(* IEC 61131-3 sources: plc-st-coding-agent/progress/evidence/f14_v10_full_20261113/jobs/custom_minimax-m27 (part 8) *)

(* ---- self-medium-01.candidate_03.st ---- *)
(* ENGINEERING_CONTRACT *)
(*
  PUB002/PUB005: valid=FALSE → loadedID:=0, valid=TRUE → loadedID:=recipe[selSlot].recipeID
  PUB006: loadCmd rising-edge triggers one-shot load; level-hold does NOT reload
  PUB007: running=TRUE blocks load, loadedID retains previous value
  PUB008: slot out-of-range [1..8] → valid=FALSE, loadedID unchanged; no array OOB access
  PUB009: validation is conjunction: recipeID<>0 AND totalRatio∈[99.0,101.0] AND temperature∈[30.0,180.0]
  Timing: state retention via VAR (static across scans); first-scan prev_* = FALSE (IEC default)
  S1: !running & rising(loadCmd) & valid-slot & empty-slot → valid=FALSE & loadedID=0
  S4/N10-S4: running → loadedID=prev(loadedID) (includes first production entry)
  N10-S9: !running & !rising(loadCmd) → both outputs retain prev value
*)
(* CONTRACT_RULES [] *)

FUNCTION_BLOCK FB
VAR_INPUT
    recipe      : ARRAY[1..8] OF ST_Recipe;
    selSlot     : INT;
    loadCmd     : BOOL;
    running     : BOOL;
END_VAR
VAR_OUTPUT
    valid       : BOOL;
    loadedID    : INT;
END_VAR
VAR
    tmp_loadTrig  : R_TRIG;
    tmp_prevRunning : BOOL := FALSE;
END_VAR

tmp_loadTrig(CLK := loadCmd);

IF tmp_loadTrig.Q AND NOT running THEN
    IF (selSlot >= 1) AND (selSlot <= 8) THEN
        IF (recipe[selSlot].recipeID <> 0) AND
           (recipe[selSlot].totalRatio >= 99.0) AND (recipe[selSlot].totalRatio <= 101.0) AND
           (recipe[selSlot].temperature >= 30.0) AND (recipe[selSlot].temperature <= 180.0) THEN
            valid    := TRUE;
            loadedID := recipe[selSlot].recipeID;
        ELSE
            valid    := FALSE;
            loadedID := 0;
        END_IF;
    ELSE
        valid    := FALSE;
    END_IF;
ELSIF running THEN
    loadedID := loadedID;
END_IF;

tmp_prevRunning := running;
END_FUNCTION_BLOCK

(* ---- self-medium-01.raw_candidate_01.st ---- *)
(* ENGINEERING_CONTRACT *)
(*
  PUB002/PUB005: valid=FALSE → loadedID:=0, valid=TRUE → loadedID:=recipe[selSlot].recipeID
  PUB006: loadCmd rising-edge triggers one-shot load; level-hold does NOT reload
  PUB007: running=TRUE blocks load, loadedID retains previous value
  PUB008: slot out-of-range [1..8] → valid=FALSE, loadedID unchanged; no array OOB access
  PUB009: validation is conjunction: recipeID<>0 AND totalRatio∈[99.0,101.0] AND temperature∈[30.0,180.0]
  Timing: state retention via VAR (static across scans); first-scan prev_* = FALSE (IEC default)
  S1: !running & rising(loadCmd) & valid-slot & empty-slot → valid=FALSE & loadedID=0
  S4/N10-S4: running → loadedID=prev(loadedID) (includes first production entry)
  N10-S9: !running & !rising(loadCmd) → both outputs retain prev value
*)
(* CONTRACT_RULES [] *)

FUNCTION_BLOCK FB
VAR_INPUT
    recipe      : ARRAY[1..8] OF ST_Recipe;
    selSlot     : INT;
    loadCmd     : BOOL;
    running     : BOOL;
END_VAR
VAR_OUTPUT
    valid       : BOOL;
    loadedID    : INT;
END_VAR
VAR
    tmp_loadTrig  : R_TRIG;
    tmp_prevRunning : BOOL := FALSE;
END_VAR

tmp_loadTrig(CLK := loadCmd);

IF tmp_loadTrig.Q AND NOT running THEN
    IF (selSlot >= 1) AND (selSlot <= 8) THEN
        IF (recipe[selSlot].recipeID <> 0) AND
           (recipe[selSlot].totalRatio >= 99.0) AND (recipe[selSlot].totalRatio <= 101.0) AND
           (recipe[selSlot].temperature >= 30.0) AND (recipe[selSlot].temperature <= 180.0) THEN
            valid    := TRUE;
            loadedID := recipe[selSlot].recipeID;
        ELSE
            valid    := FALSE;
            loadedID := 0;
        END_IF;
    ELSE
        valid    := FALSE;
    END_IF;
ELSIF running THEN
    loadedID := loadedID;
END_IF;

tmp_prevRunning := running;

(* ---- self-medium-01.raw_candidate_02.st ---- *)
(* ENGINEERING_CONTRACT *)
(*
  PUB002/PUB005: valid=FALSE → loadedID:=0, valid=TRUE → loadedID:=recipe[selSlot].recipeID
  PUB006: loadCmd rising-edge triggers one-shot load; level-hold does NOT reload
  PUB007: running=TRUE blocks load, loadedID retains previous value
  PUB008: slot out-of-range [1..8] → valid=FALSE, loadedID unchanged; no array OOB access
  PUB009: validation is conjunction: recipeID<>0 AND totalRatio∈[99.0,101.0] AND temperature∈[30.0,180.0]
  Timing: state retention via VAR (static across scans); first-scan prev_* = FALSE (IEC default)
  S1: !running & rising(loadCmd) & valid-slot & empty-slot → valid=FALSE & loadedID=0
  S4/N10-S4: running → loadedID=prev(loadedID) (includes first production entry)
  N10-S9: !running & !rising(loadCmd) → both outputs retain prev value
*)
(* CONTRACT_RULES [] *)

FUNCTION_BLOCK FB
VAR_INPUT
    recipe      : ARRAY[1..8] OF ST_Recipe;
    selSlot     : INT;
    loadCmd     : BOOL;
    running     : BOOL;
END_VAR
VAR_OUTPUT
    valid       : BOOL;
    loadedID    : INT;
END_VAR
VAR
    tmp_loadTrig  : R_TRIG;
    tmp_prevRunning : BOOL := FALSE;
END_VAR

tmp_loadTrig(CLK := loadCmd);

IF tmp_loadTrig.Q AND NOT running THEN
    IF (selSlot >= 1) AND (selSlot <= 8) THEN
        IF (recipe[selSlot].recipeID <> 0) AND
           (recipe[selSlot].totalRatio >= 99.0) AND (recipe[selSlot].totalRatio <= 101.0) AND
           (recipe[selSlot].temperature >= 30.0) AND (recipe[selSlot].temperature <= 180.0) THEN
            valid    := TRUE;
            loadedID := recipe[selSlot].recipeID;
        ELSE
            valid    := FALSE;
            loadedID := 0;
        END_IF;
    ELSE
        valid    := FALSE;
    END_IF;
ELSIF running THEN
    loadedID := loadedID;
END_IF;

tmp_prevRunning := running;
END_FUNCTION_BLOCK

(* ---- self-medium-01.raw_candidate_03.st ---- *)
(* ENGINEERING_CONTRACT *)
(*
  PUB002/PUB005: valid=FALSE → loadedID:=0, valid=TRUE → loadedID:=recipe[selSlot].recipeID
  PUB006: loadCmd rising-edge triggers one-shot load; level-hold does NOT reload
  PUB007: running=TRUE blocks load, loadedID retains previous value
  PUB008: slot out-of-range [1..8] → valid=FALSE, loadedID unchanged; no array OOB access
  PUB009: validation is conjunction: recipeID<>0 AND totalRatio∈[99.0,101.0] AND temperature∈[30.0,180.0]
  Timing: state retention via VAR (static across scans); first-scan prev_* = FALSE (IEC default)
  S1: !running & rising(loadCmd) & valid-slot & empty-slot → valid=FALSE & loadedID=0
  S4/N10-S4: running → loadedID=prev(loadedID) (includes first production entry)
  N10-S9: !running & !rising(loadCmd) → both outputs retain prev value
*)
(* CONTRACT_RULES [] *)

FUNCTION_BLOCK FB
VAR_INPUT
    recipe      : ARRAY[1..8] OF ST_Recipe;
    selSlot     : INT;
    loadCmd     : BOOL;
    running     : BOOL;
END_VAR
VAR_OUTPUT
    valid       : BOOL;
    loadedID    : INT;
END_VAR
VAR
    tmp_loadTrig  : R_TRIG;
    tmp_prevRunning : BOOL := FALSE;
END_VAR

tmp_loadTrig(CLK := loadCmd);

IF tmp_loadTrig.Q AND NOT running THEN
    IF (selSlot >= 1) AND (selSlot <= 8) THEN
        IF (recipe[selSlot].recipeID <> 0) AND
           (recipe[selSlot].totalRatio >= 99.0) AND (recipe[selSlot].totalRatio <= 101.0) AND
           (recipe[selSlot].temperature >= 30.0) AND (recipe[selSlot].temperature <= 180.0) THEN
            valid    := TRUE;
            loadedID := recipe[selSlot].recipeID;
        ELSE
            valid    := FALSE;
            loadedID := 0;
        END_IF;
    ELSE
        valid    := FALSE;
    END_IF;
ELSIF running THEN
    loadedID := loadedID;
END_IF;

tmp_prevRunning := running;
END_FUNCTION_BLOCK

(* ---- self-medium-02.candidate_01.st ---- *)
FUNCTION_BLOCK FB
VAR_INPUT
    enable     : BOOL;
    rawValue   : REAL;
END_VAR
VAR_OUTPUT
    filteredValue : REAL;
    windowFull    : BOOL;
    sampleCount   : INT;
END_VAR
VAR
    buffer     : ARRAY[0..7] OF REAL;
    writeIdx   : INT := 0;
    tmp_sum    : REAL;
    tmp_i      : INT;
END_VAR
VAR_INPUT
END_VAR
VAR_OUTPUT
END_VAR
VAR
END_VAR
(* ENGINEERING_CONTRACT
   PUB.001-004   : inputs enable, rawValue; outputs filteredValue, windowFull, sampleCount
   PUB.005       : enable=TRUE per scan: push rawValue into 8-slot ring buffer
   PUB.006       : filteredValue = mean of actually-filled slots (no zero-fill)
   PUB.007       : on windowFull: FIFO eviction of oldest sample on each new push
   PUB.008       : sampleCount = current valid samples 0..8
   PUB.009       : windowFull = TRUE when sampleCount == 8, retains TRUE thereafter
   PUB.010       : enable=FALSE: clear buffer (sampleCount=0, windowFull=FALSE),
                   filteredValue RETAINED (last computed value held)
   PUB.011       : new enable period restarts count from 1 independently
   PUB.012-015   : formal properties S1-S7 encoded as LTL constraints
   PUB.016-038   : interface unchanged; no hidden timers or global variables

   Output retention table:
   | output        | activation             | retention      | reset                    |
   |---------------|------------------------|----------------|--------------------------|
   | filteredValue | every enabled scan     | holds on FALSE | not reset; retains last  |
   | sampleCount   | increments on each push| capped at 8    | forced 0 on enable=FALSE |
   | windowFull    | set TRUE at count=8    | holds TRUE     | forced FALSE on enable=FALSE|

   Same-scan priority: disable branch executes first; rising-edge start is
   indistinguishable from normal enabled scan since buffer is pre-cleared.
   Units: filteredValue REAL; sampleCount INT 0..8; windowFull BOOL.

   CONTRACT_RULES []
*)
tmp_sum := 0.0;
IF NOT enable THEN
    sampleCount   := 0;
    windowFull    := FALSE;
    writeIdx      := 0;
ELSE
    // Push current rawValue into ring buffer
    buffer[writeIdx] := rawValue;

    // Advance write pointer (mod 8), but sampleCount only increments up to 8
    writeIdx := (writeIdx + 1) MOD 8;
    IF sampleCount < 8 THEN
        sampleCount := sampleCount + 1;
    END_IF;

    // windowFull stays TRUE once set; set it only when count reaches 8
    IF sampleCount = 8 THEN
        windowFull := TRUE;
    END_IF;

    // Compute arithmetic mean of all valid samples currently in buffer
    tmp_sum := 0.0;
    FOR tmp_i := 0 TO sampleCount - 1 DO
        tmp_sum := tmp_sum + buffer[tmp_i];
    END_FOR;
    filteredValue := tmp_sum / TO_REAL(sampleCount);
END_IF;
END_FUNCTION_BLOCK

(* ---- self-medium-02.raw_candidate_01.st ---- *)
FUNCTION_BLOCK FB
VAR_INPUT
    enable     : BOOL;
    rawValue   : REAL;
END_VAR
VAR_OUTPUT
    filteredValue : REAL;
    windowFull    : BOOL;
    sampleCount   : INT;
END_VAR
VAR
    buffer     : ARRAY[0..7] OF REAL;
    writeIdx   : INT := 0;
    tmp_sum    : REAL;
    tmp_i      : INT;
END_VAR
VAR_INPUT
END_VAR
VAR_OUTPUT
END_VAR
VAR
END_VAR
(* ENGINEERING_CONTRACT
   PUB.001-004   : inputs enable, rawValue; outputs filteredValue, windowFull, sampleCount
   PUB.005       : enable=TRUE per scan: push rawValue into 8-slot ring buffer
   PUB.006       : filteredValue = mean of actually-filled slots (no zero-fill)
   PUB.007       : on windowFull: FIFO eviction of oldest sample on each new push
   PUB.008       : sampleCount = current valid samples 0..8
   PUB.009       : windowFull = TRUE when sampleCount == 8, retains TRUE thereafter
   PUB.010       : enable=FALSE: clear buffer (sampleCount=0, windowFull=FALSE),
                   filteredValue RETAINED (last computed value held)
   PUB.011       : new enable period restarts count from 1 independently
   PUB.012-015   : formal properties S1-S7 encoded as LTL constraints
   PUB.016-038   : interface unchanged; no hidden timers or global variables

   Output retention table:
   | output        | activation             | retention      | reset                    |
   |---------------|------------------------|----------------|--------------------------|
   | filteredValue | every enabled scan     | holds on FALSE | not reset; retains last  |
   | sampleCount   | increments on each push| capped at 8    | forced 0 on enable=FALSE |
   | windowFull    | set TRUE at count=8    | holds TRUE     | forced FALSE on enable=FALSE|

   Same-scan priority: disable branch executes first; rising-edge start is
   indistinguishable from normal enabled scan since buffer is pre-cleared.
   Units: filteredValue REAL; sampleCount INT 0..8; windowFull BOOL.

   CONTRACT_RULES []
*)
tmp_sum := 0.0;
IF NOT enable THEN
    sampleCount   := 0;
    windowFull    := FALSE;
    writeIdx      := 0;
ELSE
    // Push current rawValue into ring buffer
    buffer[writeIdx] := rawValue;

    // Advance write pointer (mod 8), but sampleCount only increments up to 8
    writeIdx := (writeIdx + 1) MOD 8;
    IF sampleCount < 8 THEN
        sampleCount := sampleCount + 1;
    END_IF;

    // windowFull stays TRUE once set; set it only when count reaches 8
    IF sampleCount = 8 THEN
        windowFull := TRUE;
    END_IF;

    // Compute arithmetic mean of all valid samples currently in buffer
    tmp_sum := 0.0;
    FOR tmp_i := 0 TO sampleCount - 1 DO
        tmp_sum := tmp_sum + buffer[tmp_i];
    END_FOR;
    filteredValue := tmp_sum / TO_REAL(sampleCount);
END_IF;
END_FUNCTION_BLOCK

(* ---- self-medium-03.candidate_01.st ---- *)
(* ENGINEERING_CONTRACT *)
(*
  Gate FSM: 4 states (IDLE/OPENING/CLOSING/FAULT), obstacle safety interlock.

  PUB001: IDLE at power-on, initial button values FALSE.
  PUB003: Rising edge of openBtn (closeBtn=FALSE, openLimit=FALSE) starts opening.
          Rising edge of closeBtn (openBtn=FALSE, closeLimit=FALSE) starts closing.
          Both buttons simultaneous → no start. Commands issued same scan.
  PUB004: Buttons ignored during OPENING/CLOSING.
  PUB005: At own-direction limit → stop that direction, return IDLE.
          Opposite limit does not affect current motion.
  PUB006: MotorUp and motorDown always mutually exclusive.
  PUB007: Obstacle at any time → stop both motors, enter FAULT, errorFlag:=TRUE immediately.
          Obstacle priority > limit/motion/reset.
  PUB008: FAULT latches errorFlag, stops motors.
  PUB009: Clear fault only when: no obstacle AND both buttons new rising edge from
          not-both-pressed state to both-pressed state. Holding both with obstacle
          present does NOT clear on obstacle-clear scan. Reset→IDLE, both motors stop
          that scan, then normal PUB003 rules apply.
*)
TYPE GateState :
(
    IDLE    := 0,
    OPENING := 1,
    CLOSING := 2,
    FAULT   := 3
);
END_TYPE;

FUNCTION_BLOCK FB
VAR_INPUT
    openBtn    : BOOL;
    closeBtn   : BOOL;
    openLimit  : BOOL;
    closeLimit : BOOL;
    obstacle   : BOOL;
END_VAR

VAR_OUTPUT
    motorUp    : BOOL;
    motorDown  : BOOL;
    errorFlag  : BOOL;
END_VAR

VAR
    state        : GateState := IDLE;
    prevOpenBtn  : BOOL := FALSE;
    prevCloseBtn : BOOL := FALSE;
    prevObstacle : BOOL := FALSE;
    prevMotorUp  : BOOL := FALSE;
    prevMotorDown: BOOL := FALSE;
    prevErrorFlag: BOOL := FALSE;
END_VAR

VAR
    risingOpen  : BOOL;
    risingClose : BOOL;
    risingBoth  : BOOL;
END_VAR
(* ENGINEERING_CONTRACT *)
(*
  Gate FSM: 4 states (IDLE/OPENING/CLOSING/FAULT), obstacle safety interlock.

  PUB001: IDLE at power-on, initial button values FALSE.
  PUB003: Rising edge of openBtn (closeBtn=FALSE, openLimit=FALSE) starts opening.
          Rising edge of closeBtn (openBtn=FALSE, closeLimit=FALSE) starts closing.
          Both buttons simultaneous → no start. Commands issued same scan.
  PUB004: Buttons ignored during OPENING/CLOSING.
  PUB005: At own-direction limit → stop that direction, return IDLE.
          Opposite limit does not affect current motion.
  PUB006: MotorUp and motorDown always mutually exclusive.
  PUB007: Obstacle at any time → stop both motors, enter FAULT, errorFlag:=TRUE immediately.
          Obstacle priority > limit/motion/reset.
  PUB008: FAULT latches errorFlag, stops motors.
  PUB009: Clear fault only when: no obstacle AND both buttons new rising edge from
          not-both-pressed state to both-pressed state. Holding both with obstacle
          present does NOT clear on obstacle-clear scan. Reset→IDLE, both motors stop
          that scan, then normal PUB003 rules apply.
*)

risingOpen  := openBtn  AND NOT prevOpenBtn;
risingClose := closeBtn AND NOT prevCloseBtn;
risingBoth  := risingOpen AND risingClose;

IF obstacle THEN
    errorFlag  := TRUE;
    motorUp    := FALSE;
    motorDown  := FALSE;
    state      := FAULT;
    GOTO update_state;
END_IF;

IF state = FAULT THEN
    motorUp   := FALSE;
    motorDown := FALSE;
    IF risingBoth THEN
        errorFlag := FALSE;
        state     := IDLE;
    END_IF;
    GOTO update_state;
END_IF;

IF state = IDLE THEN
    IF risingOpen AND NOT closeBtn AND NOT openLimit THEN
        state := OPENING;
    ELSIF risingClose AND NOT openBtn AND NOT closeLimit THEN
        state := CLOSING;
    END_IF;
END_IF;

IF state = OPENING THEN
    motorUp   := TRUE;
    motorDown := FALSE;
    IF openLimit THEN
        motorUp := FALSE;
        state   := IDLE;
    END_IF;
END_IF;

IF state = CLOSING THEN
    motorUp   := FALSE;
    motorDown := TRUE;
    IF closeLimit THEN
        motorDown := FALSE;
        state     := IDLE;
    END_IF;
END_IF;

update_state:
prevOpenBtn   := openBtn;
prevCloseBtn  := closeBtn;
prevObstacle  := obstacle;
prevMotorUp   := motorUp;
prevMotorDown := motorDown;
prevErrorFlag := errorFlag;
END_FUNCTION_BLOCK
(* CONTRACT_RULES [] *)

(* ---- self-medium-03.candidate_02.st ---- *)
(* ENGINEERING_CONTRACT *)
(*
  Gate FSM: 4 states (IDLE/OPENING/CLOSING/FAULT), obstacle safety interlock.
  Priority order (highest first):
  1. Obstacle → stop both, enter FAULT, set errorFlag (same scan).
  2. FAULT → motors held FALSE; reset only on risingBoth when !obstacle.
  3. OPENING/CLOSING → motors set by state; own-limit stops and returns IDLE.
  4. IDLE → rising edge start on single valid button; simultaneous → no start.
  Motors always mutually exclusive (only one direction active at a time).
  Latched outputs: errorFlag (hold_until_reset via risingBoth).
*)
TYPE GateState :
(
    IDLE    := 0,
    OPENING := 1,
    CLOSING := 2,
    FAULT   := 3
);
END_TYPE;

FUNCTION_BLOCK FB
VAR_INPUT
    openBtn    : BOOL;
    closeBtn   : BOOL;
    openLimit  : BOOL;
    closeLimit : BOOL;
    obstacle   : BOOL;
END_VAR

VAR_OUTPUT
    motorUp    : BOOL;
    motorDown  : BOOL;
    errorFlag  : BOOL;
END_VAR

VAR
    state         : GateState := IDLE;
    prevOpenBtn   : BOOL := FALSE;
    prevCloseBtn  : BOOL := FALSE;
    prevMotorUp   : BOOL := FALSE;
    prevMotorDown : BOOL := FALSE;
    prevErrorFlag : BOOL := FALSE;
END_VAR

VAR
    risingOpen  : BOOL;
    risingClose : BOOL;
    risingBoth  : BOOL;
END_VAR

risingOpen  := openBtn  AND NOT prevOpenBtn;
risingClose := closeBtn AND NOT prevCloseBtn;
risingBoth  := openBtn AND closeBtn AND NOT prevOpenBtn AND NOT prevCloseBtn;

IF obstacle THEN
    motorUp   := FALSE;
    motorDown := FALSE;
    errorFlag := TRUE;
    state     := FAULT;
ELSE
    errorFlag := FALSE;

    IF state = FAULT THEN
        motorUp   := FALSE;
        motorDown := FALSE;
        IF risingBoth THEN
            state := IDLE;
        END_IF;

    ELSIF state = IDLE THEN
        motorUp   := FALSE;
        motorDown := FALSE;
        IF risingOpen AND NOT closeBtn AND NOT openLimit THEN
            state := OPENING;
        ELSIF risingClose AND NOT openBtn AND NOT closeLimit THEN
            state := CLOSING;
        END_IF;

    ELSIF state = OPENING THEN
        motorUp   := TRUE;
        motorDown := FALSE;
        IF openLimit THEN
            motorUp := FALSE;
            state   := IDLE;
        END_IF;

    ELSIF state = CLOSING THEN
        motorUp   := FALSE;
        motorDown := TRUE;
        IF closeLimit THEN
            motorDown := FALSE;
            state     := IDLE;
        END_IF;
    END_IF;
END_IF;

prevOpenBtn   := openBtn;
prevCloseBtn  := closeBtn;
prevMotorUp   := motorUp;
prevMotorDown := motorDown;
prevErrorFlag := errorFlag;
END_FUNCTION_BLOCK
(* CONTRACT_RULES [] *)

(* ---- self-medium-03.candidate_03.st ---- *)
Looking at the functional failures, the issue is clear from the replay: `motorUp` is not being set in the same scan as the rising edge triggers the state transition. The motor assignments need to occur after all state transitions, not interleaved within each branch.

```st
(* ENGINEERING_CONTRACT *)
(*
  Gate FSM: 4 states (IDLE/OPENING/CLOSING/FAULT), obstacle safety interlock.
  Priority order (highest first):
  1. Obstacle → stop both, enter FAULT, set errorFlag (same scan).
  2. FAULT → motors held FALSE; reset only on risingBoth when !obstacle.
  3. OPENING/CLOSING → motors set by state; own-limit stops and returns IDLE.
  4. IDLE → rising edge start on single valid button; simultaneous → no start.
  Motors always mutually exclusive (only one direction active at a time).
  Latched outputs: errorFlag (hold_until_reset via risingBoth).
*)

FUNCTION_BLOCK FB
VAR_INPUT
    openBtn    : BOOL;
    closeBtn   : BOOL;
    openLimit  : BOOL;
    closeLimit : BOOL;
    obstacle   : BOOL;
END_VAR

VAR_OUTPUT
    motorUp    : BOOL;
    motorDown  : BOOL;
    errorFlag  : BOOL;
END_VAR

VAR
    state         : INT := 0;
    prevOpenBtn   : BOOL := FALSE;
    prevCloseBtn  : BOOL := FALSE;
END_VAR

VAR
    risingOpen  : BOOL;
    risingClose : BOOL;
    risingBoth  : BOOL;
END_VAR

risingOpen  := openBtn  AND NOT prevOpenBtn;
risingClose := closeBtn AND NOT prevCloseBtn;
risingBoth  := openBtn AND closeBtn AND NOT prevOpenBtn AND NOT prevCloseBtn;

IF obstacle THEN
    state     := 3;
    errorFlag := TRUE;
ELSE
    errorFlag := FALSE;

    IF state = 3 THEN
        IF risingBoth THEN
            state := 0;
        END_IF;

    ELSIF state = 0 THEN
        IF risingOpen AND NOT closeBtn AND NOT openLimit THEN
            state := 1;
        ELSIF risingClose AND NOT openBtn AND NOT closeLimit THEN
            state := 2;
        END_IF;

    ELSIF state = 1 THEN
        IF openLimit THEN
            state := 0;
        END_IF;

    ELSIF state = 2 THEN
        IF closeLimit THEN
            state := 0;
        END_IF;
    END_IF;
END_IF;

CASE state OF
    0: motorUp := FALSE; motorDown := FALSE;
    1: motorUp := TRUE;  motorDown := FALSE;
    2: motorUp := FALSE; motorDown := TRUE;
    3: motorUp := FALSE; motorDown := FALSE;
END_CASE;

prevOpenBtn  := openBtn;
prevCloseBtn := closeBtn;
END_FUNCTION_BLOCK
(* CONTRACT_RULES [] *)

(* ---- self-medium-03.raw_candidate_01.st ---- *)
(* ENGINEERING_CONTRACT *)
(*
  Gate FSM: 4 states (IDLE/OPENING/CLOSING/FAULT), obstacle safety interlock.

  PUB001: IDLE at power-on, initial button values FALSE.
  PUB003: Rising edge of openBtn (closeBtn=FALSE, openLimit=FALSE) starts opening.
          Rising edge of closeBtn (openBtn=FALSE, closeLimit=FALSE) starts closing.
          Both buttons simultaneous → no start. Commands issued same scan.
  PUB004: Buttons ignored during OPENING/CLOSING.
  PUB005: At own-direction limit → stop that direction, return IDLE.
          Opposite limit does not affect current motion.
  PUB006: MotorUp and motorDown always mutually exclusive.
  PUB007: Obstacle at any time → stop both motors, enter FAULT, errorFlag:=TRUE immediately.
          Obstacle priority > limit/motion/reset.
  PUB008: FAULT latches errorFlag, stops motors.
  PUB009: Clear fault only when: no obstacle AND both buttons new rising edge from
          not-both-pressed state to both-pressed state. Holding both with obstacle
          present does NOT clear on obstacle-clear scan. Reset→IDLE, both motors stop
          that scan, then normal PUB003 rules apply.
*)
TYPE GateState :
(
    IDLE    := 0,
    OPENING := 1,
    CLOSING := 2,
    FAULT   := 3
);
END_TYPE

FUNCTION_BLOCK FB
VAR_INPUT
    openBtn    : BOOL;
    closeBtn   : BOOL;
    openLimit  : BOOL;
    closeLimit : BOOL;
    obstacle   : BOOL;
END_VAR

VAR_OUTPUT
    motorUp    : BOOL;
    motorDown  : BOOL;
    errorFlag  : BOOL;
END_VAR

VAR
    state        : GateState := IDLE;
    prevOpenBtn  : BOOL := FALSE;
    prevCloseBtn : BOOL := FALSE;
    prevObstacle : BOOL := FALSE;
    prevMotorUp  : BOOL := FALSE;
    prevMotorDown: BOOL := FALSE;
    prevErrorFlag: BOOL := FALSE;
END_VAR

VAR
    risingOpen  : BOOL;
    risingClose : BOOL;
    risingBoth  : BOOL;
END_VAR
(* ENGINEERING_CONTRACT *)
(*
  Gate FSM: 4 states (IDLE/OPENING/CLOSING/FAULT), obstacle safety interlock.

  PUB001: IDLE at power-on, initial button values FALSE.
  PUB003: Rising edge of openBtn (closeBtn=FALSE, openLimit=FALSE) starts opening.
          Rising edge of closeBtn (openBtn=FALSE, closeLimit=FALSE) starts closing.
          Both buttons simultaneous → no start. Commands issued same scan.
  PUB004: Buttons ignored during OPENING/CLOSING.
  PUB005: At own-direction limit → stop that direction, return IDLE.
          Opposite limit does not affect current motion.
  PUB006: MotorUp and motorDown always mutually exclusive.
  PUB007: Obstacle at any time → stop both motors, enter FAULT, errorFlag:=TRUE immediately.
          Obstacle priority > limit/motion/reset.
  PUB008: FAULT latches errorFlag, stops motors.
  PUB009: Clear fault only when: no obstacle AND both buttons new rising edge from
          not-both-pressed state to both-pressed state. Holding both with obstacle
          present does NOT clear on obstacle-clear scan. Reset→IDLE, both motors stop
          that scan, then normal PUB003 rules apply.
*)

risingOpen  := openBtn  AND NOT prevOpenBtn;
risingClose := closeBtn AND NOT prevCloseBtn;
risingBoth  := risingOpen AND risingClose;

IF obstacle THEN
    errorFlag  := TRUE;
    motorUp    := FALSE;
    motorDown  := FALSE;
    state      := FAULT;
    GOTO update_state;
END_IF

IF state = FAULT THEN
    motorUp   := FALSE;
    motorDown := FALSE;
    IF risingBoth THEN
        errorFlag := FALSE;
        state     := IDLE;
    END_IF
    GOTO update_state;
END_IF

IF state = IDLE THEN
    IF risingOpen AND NOT closeBtn AND NOT openLimit THEN
        state := OPENING;
    ELSIF risingClose AND NOT openBtn AND NOT closeLimit THEN
        state := CLOSING;
    END_IF;
END_IF;

IF state = OPENING THEN
    motorUp   := TRUE;
    motorDown := FALSE;
    IF openLimit THEN
        motorUp := FALSE;
        state   := IDLE;
    END_IF;
END_IF;

IF state = CLOSING THEN
    motorUp   := FALSE;
    motorDown := TRUE;
    IF closeLimit THEN
        motorDown := FALSE;
        state     := IDLE;
    END_IF;
END_IF;

update_state:
prevOpenBtn   := openBtn;
prevCloseBtn  := closeBtn;
prevObstacle  := obstacle;
prevMotorUp   := motorUp;
prevMotorDown := motorDown;
prevErrorFlag := errorFlag;
END_FUNCTION_BLOCK
(* CONTRACT_RULES [] *)

(* ---- self-medium-03.raw_candidate_02.st ---- *)
(* ENGINEERING_CONTRACT *)
(*
  Gate FSM: 4 states (IDLE/OPENING/CLOSING/FAULT), obstacle safety interlock.
  Priority order (highest first):
  1. Obstacle → stop both, enter FAULT, set errorFlag (same scan).
  2. FAULT → motors held FALSE; reset only on risingBoth when !obstacle.
  3. OPENING/CLOSING → motors set by state; own-limit stops and returns IDLE.
  4. IDLE → rising edge start on single valid button; simultaneous → no start.
  Motors always mutually exclusive (only one direction active at a time).
  Latched outputs: errorFlag (hold_until_reset via risingBoth).
*)
TYPE GateState :
(
    IDLE    := 0,
    OPENING := 1,
    CLOSING := 2,
    FAULT   := 3
);
END_TYPE

FUNCTION_BLOCK FB
VAR_INPUT
    openBtn    : BOOL;
    closeBtn   : BOOL;
    openLimit  : BOOL;
    closeLimit : BOOL;
    obstacle   : BOOL;
END_VAR

VAR_OUTPUT
    motorUp    : BOOL;
    motorDown  : BOOL;
    errorFlag  : BOOL;
END_VAR

VAR
    state         : GateState := IDLE;
    prevOpenBtn   : BOOL := FALSE;
    prevCloseBtn  : BOOL := FALSE;
    prevMotorUp   : BOOL := FALSE;
    prevMotorDown : BOOL := FALSE;
    prevErrorFlag : BOOL := FALSE;
END_VAR

VAR
    risingOpen  : BOOL;
    risingClose : BOOL;
    risingBoth  : BOOL;
END_VAR

risingOpen  := openBtn  AND NOT prevOpenBtn;
risingClose := closeBtn AND NOT prevCloseBtn;
risingBoth  := openBtn AND closeBtn AND NOT prevOpenBtn AND NOT prevCloseBtn;

IF obstacle THEN
    motorUp   := FALSE;
    motorDown := FALSE;
    errorFlag := TRUE;
    state     := FAULT;
ELSE
    errorFlag := FALSE;

    IF state = FAULT THEN
        motorUp   := FALSE;
        motorDown := FALSE;
        IF risingBoth THEN
            state := IDLE;
        END_IF;

    ELSIF state = IDLE THEN
        motorUp   := FALSE;
        motorDown := FALSE;
        IF risingOpen AND NOT closeBtn AND NOT openLimit THEN
            state := OPENING;
        ELSIF risingClose AND NOT openBtn AND NOT closeLimit THEN
            state := CLOSING;
        END_IF;

    ELSIF state = OPENING THEN
        motorUp   := TRUE;
        motorDown := FALSE;
        IF openLimit THEN
            motorUp := FALSE;
            state   := IDLE;
        END_IF;

    ELSIF state = CLOSING THEN
        motorUp   := FALSE;
        motorDown := TRUE;
        IF closeLimit THEN
            motorDown := FALSE;
            state     := IDLE;
        END_IF;
    END_IF;
END_IF;

prevOpenBtn   := openBtn;
prevCloseBtn  := closeBtn;
prevMotorUp   := motorUp;
prevMotorDown := motorDown;
prevErrorFlag := errorFlag;
END_FUNCTION_BLOCK
(* CONTRACT_RULES [] *)

(* ---- self-medium-03.raw_candidate_03.st ---- *)
Looking at the functional failures, the issue is clear from the replay: `motorUp` is not being set in the same scan as the rising edge triggers the state transition. The motor assignments need to occur after all state transitions, not interleaved within each branch.

```st
(* ENGINEERING_CONTRACT *)
(*
  Gate FSM: 4 states (IDLE/OPENING/CLOSING/FAULT), obstacle safety interlock.
  Priority order (highest first):
  1. Obstacle → stop both, enter FAULT, set errorFlag (same scan).
  2. FAULT → motors held FALSE; reset only on risingBoth when !obstacle.
  3. OPENING/CLOSING → motors set by state; own-limit stops and returns IDLE.
  4. IDLE → rising edge start on single valid button; simultaneous → no start.
  Motors always mutually exclusive (only one direction active at a time).
  Latched outputs: errorFlag (hold_until_reset via risingBoth).
*)

FUNCTION_BLOCK FB
VAR_INPUT
    openBtn    : BOOL;
    closeBtn   : BOOL;
    openLimit  : BOOL;
    closeLimit : BOOL;
    obstacle   : BOOL;
END_VAR

VAR_OUTPUT
    motorUp    : BOOL;
    motorDown  : BOOL;
    errorFlag  : BOOL;
END_VAR

VAR
    state         : INT := 0;
    prevOpenBtn   : BOOL := FALSE;
    prevCloseBtn  : BOOL := FALSE;
END_VAR

VAR
    risingOpen  : BOOL;
    risingClose : BOOL;
    risingBoth  : BOOL;
END_VAR

risingOpen  := openBtn  AND NOT prevOpenBtn;
risingClose := closeBtn AND NOT prevCloseBtn;
risingBoth  := openBtn AND closeBtn AND NOT prevOpenBtn AND NOT prevCloseBtn;

IF obstacle THEN
    state     := 3;
    errorFlag := TRUE;
ELSE
    errorFlag := FALSE;

    IF state = 3 THEN
        IF risingBoth THEN
            state := 0;
        END_IF;

    ELSIF state = 0 THEN
        IF risingOpen AND NOT closeBtn AND NOT openLimit THEN
            state := 1;
        ELSIF risingClose AND NOT openBtn AND NOT closeLimit THEN
            state := 2;
        END_IF;

    ELSIF state = 1 THEN
        IF openLimit THEN
            state := 0;
        END_IF;

    ELSIF state = 2 THEN
        IF closeLimit THEN
            state := 0;
        END_IF;
    END_IF;
END_IF;

CASE state OF
    0: motorUp := FALSE; motorDown := FALSE;
    1: motorUp := TRUE;  motorDown := FALSE;
    2: motorUp := FALSE; motorDown := TRUE;
    3: motorUp := FALSE; motorDown := FALSE;
END_CASE;

prevOpenBtn  := openBtn;
prevCloseBtn := closeBtn;
END_FUNCTION_BLOCK
(* CONTRACT_RULES [] *)

(* ---- self-medium-04.candidate_01.st ---- *)
FUNCTION_BLOCK FB
VAR_INPUT
    startBtn    : BOOL;
    resetBtn    : BOOL;
    doneSensor  : BOOL;
    targetVol   : REAL;
    flowVol     : REAL;
END_VAR
VAR_OUTPUT
    valveOpen   : BOOL := FALSE;
    fillsToday  : INT  := 0;
END_VAR
VAR
    state           : INT := 0; // 0=IDLE, 1=FILLING, 2=WAIT_CONFIRM
    accumulated     : REAL := 0.0;
    pendingConfirm  : BOOL := FALSE;
    prevStartBtn    : BOOL := FALSE;
    prevResetBtn    : BOOL := FALSE;
    prevValveOpen   : BOOL := FALSE;
    R_TRIG_reset    : R_TRIG;
    R_TRIG_start    : R_TRIG;
END_VAR
VAR_CONSTANT
    IDLE          : INT := 0;
    FILLING       : INT := 1;
    WAIT_CONFIRM  : INT := 2;
END_VAR
BEGIN
    (* ENGINEERING_CONTRACT
    ---------------------------------------------------------------------
    PUB001: Initialization - valve closed (valveOpen=FALSE), no pending
            confirmation (pendingConfirm=FALSE), fillsToday=0 on cold start.
    PUB002: Rising-edge detection for startBtn/resetBtn; pre-power state FALSE.
    PUB003: Scan execution order: reset(1)→start/new-bottle(2)→accumulate/
            close-on-target(3)→doneSensor read→confirm/count(4).
    PUB004: resetBtn rising edge has highest priority; clears all state,
            ignores same-scan start/flow/confirmation.
    PUB005: startBtn rising edge in IDLE/WAIT_CONFIRM starts new bottle,
            clears accumulation, opens valve. Prior pendingConfirm cancelled.
            New start during FILLING does NOT reset current bottle.
    PUB006: Accumulate flowVol every scan including startup scan.
    PUB007: When accumulated >= targetVol, close valve and set pendingConfirm
            immediately in same scan.
    PUB008: After closing, read doneSensor same scan. If TRUE, confirm/count
            immediately. If FALSE, wait for first TRUE (unless reset/new-start).
    PUB009: Each confirmation increments fillsToday by 1. At 32767, confirm
            completes but count stays at 32767.
    PUB010: Confirmation clears pendingConfirm. Continuous TRUE does not
            double-count. New-bottle start-cancel clears pendingConfirm.
    PUB011: fillsToday is INT; reset clears to 0.
    ---------------------------------------------------------------------
    OUTPUT RETENTION:
    - valveOpen: held open during FILLING until target met or reset/start.
    - fillsToday: monotonic non-decreasing except reset (S3); max 32767.
    - pendingConfirm: held TRUE from close until first TRUE doneSensor.
    EXPLICIT RESET: resetBtn rising edge clears accumulated, fillsToday,
            valveOpen, pendingConfirm, state→IDLE.
    SAME-SCAN PRIORITY: reset > close-on-target-with-confirm > start.
    UNITS/BOUNDARIES: accumulated REAL mL; fillsToday INT [0..32767];
            targetVol, flowVol REAL mL.
    ---------------------------------------------------------------------
    *)

    // --- Step 1: Reset (highest priority) ---
    R_TRIG_reset(CLK := resetBtn);
    IF R_TRIG_reset.Q THEN
        accumulated    := 0.0;
        fillsToday     := 0;
        valveOpen      := FALSE;
        pendingConfirm := FALSE;
        state          := IDLE;
        GOTO end_scan;
    END_IF;

    // --- Step 2: Start new bottle ---
    R_TRIG_start(CLK := startBtn);
    IF R_TRIG_start.Q THEN
        IF state = WAIT_CONFIRM THEN
            pendingConfirm := FALSE;
        END_IF;
        IF state <> FILLING THEN
            accumulated  := 0.0;
            valveOpen    := TRUE;
            state        := FILLING;
        END_IF;
    END_IF;

    // --- Step 3: Accumulate and close on target ---
    IF state = FILLING THEN
        accumulated := accumulated + flowVol;
        IF accumulated >= targetVol THEN
            valveOpen      := FALSE;
            pendingConfirm := TRUE;
        END_IF;
    END_IF;

    // --- Step 4: Read doneSensor after close, confirm/count ---
    IF pendingConfirm THEN
        IF doneSensor THEN
            IF fillsToday < 32767 THEN
                fillsToday := fillsToday + 1;
            END_IF;
            pendingConfirm := FALSE;
            state          := IDLE;
        END_IF;
    END_IF;

    // Track valve transition for S10 (non-reset close → confirm next scan)
    // State WAIT_CONFIRM entered when valve just closed without immediate confirm
    IF prevValveOpen AND NOT valveOpen AND NOT R_TRIG_reset.Q AND state = WAIT_CONFIRM THEN
        IF doneSensor THEN
            IF fillsToday < 32767 THEN
                fillsToday := fillsToday + 1;
            END_IF;
            pendingConfirm := FALSE;
            state          := IDLE;
        END_IF;
    END_IF;

    end_scan:
    // Update previous states for edge detection
    prevStartBtn  := startBtn;
    prevResetBtn  := resetBtn;
    prevValveOpen := valveOpen;
END_FUNCTION_BLOCK

(* ---- self-medium-04.candidate_02.st ---- *)
FUNCTION_BLOCK FB
VAR_INPUT
    startBtn    : BOOL;
    resetBtn    : BOOL;
    doneSensor  : BOOL;
    targetVol   : REAL;
    flowVol     : REAL;
END_VAR
VAR_OUTPUT
    valveOpen   : BOOL := FALSE;
    fillsToday  : INT  := 0;
END_VAR
VAR
    state          : INT := 0;
    accumulated    : REAL := 0.0;
    pendingConfirm : BOOL := FALSE;
    prevStartBtn   : BOOL := FALSE;
    prevResetBtn   : BOOL := FALSE;
    prevValveOpen  : BOOL := FALSE;
END_VAR
BEGIN
    (* ENGINEERING_CONTRACT
    ---------------------------------------------------------------------
    PUB001: Initialization - valve closed (valveOpen=FALSE), no pending
            confirmation (pendingConfirm=FALSE), fillsToday=0 on cold start.
    PUB002: Rising-edge detection for startBtn/resetBtn; pre-power state FALSE.
    PUB003: Scan execution order: reset(1)→start/new-bottle(2)→accumulate/
            close-on-target(3)→doneSensor read→confirm/count(4).
    PUB004: resetBtn rising edge has highest priority; clears all state,
            ignores same-scan start/flow/confirmation.
    PUB005: startBtn rising edge in IDLE(0)/WAIT_CONFIRM(2) starts new bottle,
            clears accumulation, opens valve. Prior pendingConfirm cancelled.
            New start during FILLING(1) does NOT reset current bottle.
    PUB006: Accumulate flowVol every scan including startup scan.
    PUB007: When accumulated >= targetVol, close valve and set pendingConfirm
            immediately in same scan.
    PUB008: After closing, read doneSensor same scan. If TRUE, confirm/count
            immediately. If FALSE, wait for first TRUE (unless reset/new-start).
    PUB009: Each confirmation increments fillsToday by 1. At 32767, confirm
            completes but count stays at 32767.
    PUB010: Confirmation clears pendingConfirm. Continuous TRUE does not
            double-count. New-bottle start-cancel clears pendingConfirm.
    PUB011: fillsToday is INT; reset clears to 0.
    ---------------------------------------------------------------------
    OUTPUT RETENTION:
    - valveOpen: held open during FILLING until target met or reset/start.
    - fillsToday: monotonic non-decreasing except reset (S3); max 32767.
    - pendingConfirm: held TRUE from close until first TRUE doneSensor.
    EXPLICIT RESET: resetBtn rising edge clears accumulated, fillsToday,
            valveOpen, pendingConfirm, state→0(IDLE).
    SAME-SCAN PRIORITY: reset > close-on-target-with-confirm > start.
    UNITS/BOUNDARIES: accumulated REAL mL; fillsToday INT [0..32767];
            targetVol, flowVol REAL mL.
    ---------------------------------------------------------------------
    *)

    // --- Step 1: Reset (highest priority) ---
    IF resetBtn AND NOT prevResetBtn THEN
        accumulated    := 0.0;
        fillsToday     := 0;
        valveOpen      := FALSE;
        pendingConfirm := FALSE;
        state          := 0;
        prevStartBtn   := startBtn;
        prevResetBtn   := resetBtn;
        prevValveOpen  := FALSE;
        RETURN;
    END_IF;

    // --- Step 2: Start new bottle ---
    IF startBtn AND NOT prevStartBtn THEN
        IF state = 2 THEN
            pendingConfirm := FALSE;
        END_IF;
        IF state <> 1 THEN
            accumulated := 0.0;
            valveOpen   := TRUE;
            state       := 1;
        END_IF;
    END_IF;

    // --- Step 3: Accumulate and close on target ---
    IF state = 1 THEN
        accumulated := accumulated + flowVol;
        IF accumulated >= targetVol THEN
            valveOpen      := FALSE;
            pendingConfirm := TRUE;
            state          := 2;
        END_IF;
    END_IF;

    // --- Step 4: Read doneSensor and confirm/count ---
    IF pendingConfirm THEN
        IF doneSensor THEN
            IF fillsToday < 32767 THEN
                fillsToday := fillsToday + 1;
            END_IF;
            pendingConfirm := FALSE;
            state          := 0;
        END_IF;
    END_IF;

    // Update previous states for next scan edge detection
    prevStartBtn  := startBtn;
    prevResetBtn  := resetBtn;
    prevValveOpen := valveOpen;
END_FUNCTION_BLOCK

(* ---- self-medium-04.candidate_03.st ---- *)
FUNCTION_BLOCK FB
VAR_INPUT
    startBtn    : BOOL;
    resetBtn    : BOOL;
    doneSensor  : BOOL;
    targetVol   : REAL;
    flowVol     : REAL;
END_VAR
VAR_OUTPUT
    valveOpen   : BOOL := FALSE;
    fillsToday  : INT  := 0;
END_VAR
VAR
    state           : INT := 0; // 0=IDLE, 1=FILLING, 2=WAIT_CONFIRM
    accumulated     : REAL := 0.0;
    pendingConfirm  : BOOL := FALSE;
    prevStartBtn    : BOOL := FALSE;
    prevResetBtn    : BOOL := FALSE;
    prevValveOpen   : BOOL := FALSE;
    R_TRIG_reset    : R_TRIG;
    R_TRIG_start    : R_TRIG;
END_VAR
BEGIN
    // --- Step 1: Reset (highest priority) ---
    R_TRIG_reset(CLK := resetBtn);
    IF R_TRIG_reset.Q THEN
        accumulated    := 0.0;
        fillsToday     := 0;
        valveOpen      := FALSE;
        pendingConfirm := FALSE;
        state          := 0; // IDLE
    ELSE
        // --- Step 2: Start new bottle ---
        R_TRIG_start(CLK := startBtn);
        IF R_TRIG_start.Q THEN
            IF state = 2 THEN // WAIT_CONFIRM
                pendingConfirm := FALSE;
            END_IF;
            IF state <> 1 THEN // not FILLING
                accumulated := 0.0;
                valveOpen   := TRUE;
                state       := 1; // FILLING
            END_IF;
        END_IF;

        // --- Step 3: Accumulate and close on target ---
        IF state = 1 THEN // FILLING
            accumulated := accumulated + flowVol;
            IF accumulated >= targetVol THEN
                valveOpen      := FALSE;
                pendingConfirm := TRUE;
                state          := 2; // WAIT_CONFIRM
            END_IF;
        END_IF;

        // --- Step 4: Confirm/count (same-scan or deferred) ---
        IF prevValveOpen AND NOT valveOpen AND pendingConfirm THEN
            // Valve just closed this scan
            IF doneSensor THEN
                IF fillsToday < 32767 THEN
                    fillsToday := fillsToday + 1;
                END_IF;
                pendingConfirm := FALSE;
                state          := 0; // IDLE
            END_IF;
        ELSIF pendingConfirm AND doneSensor THEN
            // S10: Valve closed last scan, confirmed this scan
            IF fillsToday < 32767 THEN
                fillsToday := fillsToday + 1;
            END_IF;
            pendingConfirm := FALSE;
            state          := 0; // IDLE
        END_IF;
    END_IF;

    prevStartBtn  := startBtn;
    prevResetBtn  := resetBtn;
    prevValveOpen := valveOpen;
END_FUNCTION_BLOCK

(* ---- self-medium-04.candidate_04.st ---- *)
FUNCTION_BLOCK FB
VAR_INPUT
    startBtn    : BOOL;
    resetBtn    : BOOL;
    doneSensor  : BOOL;
    targetVol   : REAL;
    flowVol     : REAL;
END_VAR
VAR_OUTPUT
    valveOpen   : BOOL := FALSE;
    fillsToday  : INT  := 0;
END_VAR
VAR
    state           : INT := 0; // 0=IDLE, 1=FILLING, 2=WAIT_CONFIRM
    accumulated     : REAL := 0.0;
    pendingConfirm  : BOOL := FALSE;
    prevStartBtn    : BOOL := FALSE;
    prevResetBtn    : BOOL := FALSE;
    prevValveOpen   : BOOL := FALSE;
    R_TRIG_reset    : R_TRIG;
    R_TRIG_start    : R_TRIG;
END_VAR
BEGIN
    (* ENGINEERING_CONTRACT
    ---------------------------------------------------------------------
    PUB001: Initialization - valve closed (valveOpen=FALSE), no pending
            confirmation (pendingConfirm=FALSE), fillsToday=0 on cold start.
    PUB002: Rising-edge detection for startBtn/resetBtn; pre-power state FALSE.
    PUB003: Scan execution order: reset(1)→start/new-bottle(2)→accumulate/
            close-on-target(3)→doneSensor read→confirm/count(4).
    PUB004: resetBtn rising edge has highest priority; clears all state,
            ignores same-scan start/flow/confirmation.
    PUB005: startBtn rising edge in IDLE/WAIT_CONFIRM starts new bottle,
            clears accumulation, opens valve. Prior pendingConfirm cancelled.
            New start during FILLING does NOT reset current bottle.
    PUB006: Accumulate flowVol every scan including startup scan.
    PUB007: When accumulated >= targetVol, close valve and set pendingConfirm
            immediately in same scan.
    PUB008: After closing, read doneSensor same scan. If TRUE, confirm/count
            immediately. If FALSE, wait for first TRUE (unless reset/new-start).
    PUB009: Each confirmation increments fillsToday by 1. At 32767, confirm
            completes but count stays at 32767.
    PUB010: Confirmation clears pendingConfirm. Continuous TRUE does not
            double-count. New-bottle start-cancel clears pendingConfirm.
    PUB011: fillsToday is INT; reset clears to 0.
    ---------------------------------------------------------------------
    OUTPUT RETENTION:
    - valveOpen: held open during FILLING until target met or reset/start.
    - fillsToday: monotonic non-decreasing except reset (S3); max 32767.
    - pendingConfirm: held TRUE from close until first TRUE doneSensor.
    EXPLICIT RESET: resetBtn rising edge clears accumulated, fillsToday,
            valveOpen, pendingConfirm, state→0(IDLE).
    SAME-SCAN PRIORITY: reset > close-on-target-with-confirm > start.
    UNITS/BOUNDARIES: accumulated REAL mL; fillsToday INT [0..32767];
            targetVol, flowVol REAL mL.
    ---------------------------------------------------------------------
    *)

    // Update edge detectors every scan
    R_TRIG_reset(CLK := resetBtn);
    R_TRIG_start(CLK := startBtn);

    // --- Step 1: Reset (highest priority) ---
    IF R_TRIG_reset.Q THEN
        accumulated    := 0.0;
        fillsToday     := 0;
        valveOpen      := FALSE;
        pendingConfirm := FALSE;
        state          := 0; // IDLE
        prevValveOpen  := FALSE;
        prevStartBtn   := startBtn;
        prevResetBtn   := resetBtn;
        RETURN;
    END_IF;

    // --- Step 2: Start new bottle ---
    IF R_TRIG_start.Q THEN
        IF state = 2 THEN // WAIT_CONFIRM
            pendingConfirm := FALSE;
        END_IF;
        IF state <> 1 THEN // not FILLING
            accumulated  := 0.0;
            valveOpen    := TRUE;
            state        := 1; // FILLING
        END_IF;
    END_IF;

    // --- Step 3: Accumulate and close on target ---
    IF state = 1 THEN // FILLING
        accumulated := accumulated + flowVol;
        IF accumulated >= targetVol THEN
            valveOpen      := FALSE;
            pendingConfirm := TRUE;
            state          := 2; // WAIT_CONFIRM
        END_IF;
    END_IF;

    // --- Step 4: Confirm/count on doneSensor ---
    IF pendingConfirm THEN
        IF doneSensor THEN
            IF fillsToday < 32767 THEN
                fillsToday := fillsToday + 1;
            END_IF;
            pendingConfirm := FALSE;
            state          := 0; // IDLE
        END_IF;
    END_IF;

    // Update previous states for edge detection
    prevStartBtn  := startBtn;
    prevResetBtn  := resetBtn;
    prevValveOpen := valveOpen;
END_FUNCTION_BLOCK

(* ---- self-medium-04.raw_candidate_01.st ---- *)
FUNCTION_BLOCK FB
VAR_INPUT
    startBtn    : BOOL;
    resetBtn    : BOOL;
    doneSensor  : BOOL;
    targetVol   : REAL;
    flowVol     : REAL;
END_VAR
VAR_OUTPUT
    valveOpen   : BOOL := FALSE;
    fillsToday  : INT  := 0;
END_VAR
VAR
    state           : INT := 0; // 0=IDLE, 1=FILLING, 2=WAIT_CONFIRM
    accumulated     : REAL := 0.0;
    pendingConfirm  : BOOL := FALSE;
    prevStartBtn    : BOOL := FALSE;
    prevResetBtn    : BOOL := FALSE;
    prevValveOpen   : BOOL := FALSE;
    R_TRIG_reset    : R_TRIG;
    R_TRIG_start    : R_TRIG;
END_VAR
VAR_CONSTANT
    IDLE          : INT := 0;
    FILLING       : INT := 1;
    WAIT_CONFIRM  : INT := 2;
END_VAR
BEGIN
    (* ENGINEERING_CONTRACT
    ---------------------------------------------------------------------
    PUB001: Initialization - valve closed (valveOpen=FALSE), no pending
            confirmation (pendingConfirm=FALSE), fillsToday=0 on cold start.
    PUB002: Rising-edge detection for startBtn/resetBtn; pre-power state FALSE.
    PUB003: Scan execution order: reset(1)→start/new-bottle(2)→accumulate/
            close-on-target(3)→doneSensor read→confirm/count(4).
    PUB004: resetBtn rising edge has highest priority; clears all state,
            ignores same-scan start/flow/confirmation.
    PUB005: startBtn rising edge in IDLE/WAIT_CONFIRM starts new bottle,
            clears accumulation, opens valve. Prior pendingConfirm cancelled.
            New start during FILLING does NOT reset current bottle.
    PUB006: Accumulate flowVol every scan including startup scan.
    PUB007: When accumulated >= targetVol, close valve and set pendingConfirm
            immediately in same scan.
    PUB008: After closing, read doneSensor same scan. If TRUE, confirm/count
            immediately. If FALSE, wait for first TRUE (unless reset/new-start).
    PUB009: Each confirmation increments fillsToday by 1. At 32767, confirm
            completes but count stays at 32767.
    PUB010: Confirmation clears pendingConfirm. Continuous TRUE does not
            double-count. New-bottle start-cancel clears pendingConfirm.
    PUB011: fillsToday is INT; reset clears to 0.
    ---------------------------------------------------------------------
    OUTPUT RETENTION:
    - valveOpen: held open during FILLING until target met or reset/start.
    - fillsToday: monotonic non-decreasing except reset (S3); max 32767.
    - pendingConfirm: held TRUE from close until first TRUE doneSensor.
    EXPLICIT RESET: resetBtn rising edge clears accumulated, fillsToday,
            valveOpen, pendingConfirm, state→IDLE.
    SAME-SCAN PRIORITY: reset > close-on-target-with-confirm > start.
    UNITS/BOUNDARIES: accumulated REAL mL; fillsToday INT [0..32767];
            targetVol, flowVol REAL mL.
    ---------------------------------------------------------------------
    *)

    // --- Step 1: Reset (highest priority) ---
    R_TRIG_reset(CLK := resetBtn);
    IF R_TRIG_reset.Q THEN
        accumulated    := 0.0;
        fillsToday     := 0;
        valveOpen      := FALSE;
        pendingConfirm := FALSE;
        state          := IDLE;
        GOTO end_scan;
    END_IF

    // --- Step 2: Start new bottle ---
    R_TRIG_start(CLK := startBtn);
    IF R_TRIG_start.Q THEN
        IF state = WAIT_CONFIRM THEN
            pendingConfirm := FALSE;
        END_IF
        IF state <> FILLING THEN
            accumulated  := 0.0;
            valveOpen    := TRUE;
            state        := FILLING;
        END_IF;
    END_IF

    // --- Step 3: Accumulate and close on target ---
    IF state = FILLING THEN
        accumulated := accumulated + flowVol;
        IF accumulated >= targetVol THEN
            valveOpen      := FALSE;
            pendingConfirm := TRUE;
        END_IF;
    END_IF

    // --- Step 4: Read doneSensor after close, confirm/count ---
    IF pendingConfirm THEN
        IF doneSensor THEN
            IF fillsToday < 32767 THEN
                fillsToday := fillsToday + 1;
            END_IF;
            pendingConfirm := FALSE;
            state          := IDLE;
        END_IF;
    END_IF

    // Track valve transition for S10 (non-reset close → confirm next scan)
    // State WAIT_CONFIRM entered when valve just closed without immediate confirm
    IF prevValveOpen AND NOT valveOpen AND NOT R_TRIG_reset.Q AND state = WAIT_CONFIRM THEN
        IF doneSensor THEN
            IF fillsToday < 32767 THEN
                fillsToday := fillsToday + 1;
            END_IF;
            pendingConfirm := FALSE;
            state          := IDLE;
        END_IF;
    END_IF;

    end_scan:
    // Update previous states for edge detection
    prevStartBtn  := startBtn;
    prevResetBtn  := resetBtn;
    prevValveOpen := valveOpen;
END_FUNCTION_BLOCK

(* ---- self-medium-04.raw_candidate_02.st ---- *)
FUNCTION_BLOCK FB
VAR_INPUT
    startBtn    : BOOL;
    resetBtn    : BOOL;
    doneSensor  : BOOL;
    targetVol   : REAL;
    flowVol     : REAL;
END_VAR
VAR_OUTPUT
    valveOpen   : BOOL := FALSE;
    fillsToday  : INT  := 0;
END_VAR
VAR
    state          : INT := 0;
    accumulated    : REAL := 0.0;
    pendingConfirm : BOOL := FALSE;
    prevStartBtn   : BOOL := FALSE;
    prevResetBtn   : BOOL := FALSE;
    prevValveOpen  : BOOL := FALSE;
END_VAR
BEGIN
    (* ENGINEERING_CONTRACT
    ---------------------------------------------------------------------
    PUB001: Initialization - valve closed (valveOpen=FALSE), no pending
            confirmation (pendingConfirm=FALSE), fillsToday=0 on cold start.
    PUB002: Rising-edge detection for startBtn/resetBtn; pre-power state FALSE.
    PUB003: Scan execution order: reset(1)→start/new-bottle(2)→accumulate/
            close-on-target(3)→doneSensor read→confirm/count(4).
    PUB004: resetBtn rising edge has highest priority; clears all state,
            ignores same-scan start/flow/confirmation.
    PUB005: startBtn rising edge in IDLE(0)/WAIT_CONFIRM(2) starts new bottle,
            clears accumulation, opens valve. Prior pendingConfirm cancelled.
            New start during FILLING(1) does NOT reset current bottle.
    PUB006: Accumulate flowVol every scan including startup scan.
    PUB007: When accumulated >= targetVol, close valve and set pendingConfirm
            immediately in same scan.
    PUB008: After closing, read doneSensor same scan. If TRUE, confirm/count
            immediately. If FALSE, wait for first TRUE (unless reset/new-start).
    PUB009: Each confirmation increments fillsToday by 1. At 32767, confirm
            completes but count stays at 32767.
    PUB010: Confirmation clears pendingConfirm. Continuous TRUE does not
            double-count. New-bottle start-cancel clears pendingConfirm.
    PUB011: fillsToday is INT; reset clears to 0.
    ---------------------------------------------------------------------
    OUTPUT RETENTION:
    - valveOpen: held open during FILLING until target met or reset/start.
    - fillsToday: monotonic non-decreasing except reset (S3); max 32767.
    - pendingConfirm: held TRUE from close until first TRUE doneSensor.
    EXPLICIT RESET: resetBtn rising edge clears accumulated, fillsToday,
            valveOpen, pendingConfirm, state→0(IDLE).
    SAME-SCAN PRIORITY: reset > close-on-target-with-confirm > start.
    UNITS/BOUNDARIES: accumulated REAL mL; fillsToday INT [0..32767];
            targetVol, flowVol REAL mL.
    ---------------------------------------------------------------------
    *)

    // --- Step 1: Reset (highest priority) ---
    IF resetBtn AND NOT prevResetBtn THEN
        accumulated    := 0.0;
        fillsToday     := 0;
        valveOpen      := FALSE;
        pendingConfirm := FALSE;
        state          := 0;
        prevStartBtn   := startBtn;
        prevResetBtn   := resetBtn;
        prevValveOpen  := FALSE;
        RETURN;
    END_IF;

    // --- Step 2: Start new bottle ---
    IF startBtn AND NOT prevStartBtn THEN
        IF state = 2 THEN
            pendingConfirm := FALSE;
        END_IF;
        IF state <> 1 THEN
            accumulated := 0.0;
            valveOpen   := TRUE;
            state       := 1;
        END_IF;
    END_IF;

    // --- Step 3: Accumulate and close on target ---
    IF state = 1 THEN
        accumulated := accumulated + flowVol;
        IF accumulated >= targetVol THEN
            valveOpen      := FALSE;
            pendingConfirm := TRUE;
            state          := 2;
        END_IF;
    END_IF;

    // --- Step 4: Read doneSensor and confirm/count ---
    IF pendingConfirm THEN
        IF doneSensor THEN
            IF fillsToday < 32767 THEN
                fillsToday := fillsToday + 1;
            END_IF;
            pendingConfirm := FALSE;
            state          := 0;
        END_IF;
    END_IF;

    // Update previous states for next scan edge detection
    prevStartBtn  := startBtn;
    prevResetBtn  := resetBtn;
    prevValveOpen := valveOpen;
END_FUNCTION_BLOCK

(* ---- self-medium-04.raw_candidate_03.st ---- *)
FUNCTION_BLOCK FB
VAR_INPUT
    startBtn    : BOOL;
    resetBtn    : BOOL;
    doneSensor  : BOOL;
    targetVol   : REAL;
    flowVol     : REAL;
END_VAR
VAR_OUTPUT
    valveOpen   : BOOL := FALSE;
    fillsToday  : INT  := 0;
END_VAR
VAR
    state           : INT := 0; // 0=IDLE, 1=FILLING, 2=WAIT_CONFIRM
    accumulated     : REAL := 0.0;
    pendingConfirm  : BOOL := FALSE;
    prevStartBtn    : BOOL := FALSE;
    prevResetBtn    : BOOL := FALSE;
    prevValveOpen   : BOOL := FALSE;
    R_TRIG_reset    : R_TRIG;
    R_TRIG_start    : R_TRIG;
END_VAR
BEGIN
    // --- Step 1: Reset (highest priority) ---
    R_TRIG_reset(CLK := resetBtn);
    IF R_TRIG_reset.Q THEN
        accumulated    := 0.0;
        fillsToday     := 0;
        valveOpen      := FALSE;
        pendingConfirm := FALSE;
        state          := 0; // IDLE
    ELSE
        // --- Step 2: Start new bottle ---
        R_TRIG_start(CLK := startBtn);
        IF R_TRIG_start.Q THEN
            IF state = 2 THEN // WAIT_CONFIRM
                pendingConfirm := FALSE;
            END_IF;
            IF state <> 1 THEN // not FILLING
                accumulated := 0.0;
                valveOpen   := TRUE;
                state       := 1; // FILLING
            END_IF;
        END_IF;

        // --- Step 3: Accumulate and close on target ---
        IF state = 1 THEN // FILLING
            accumulated := accumulated + flowVol;
            IF accumulated >= targetVol THEN
                valveOpen      := FALSE;
                pendingConfirm := TRUE;
                state          := 2; // WAIT_CONFIRM
            END_IF;
        END_IF;

        // --- Step 4: Confirm/count (same-scan or deferred) ---
        IF prevValveOpen AND NOT valveOpen AND pendingConfirm THEN
            // Valve just closed this scan
            IF doneSensor THEN
                IF fillsToday < 32767 THEN
                    fillsToday := fillsToday + 1;
                END_IF;
                pendingConfirm := FALSE;
                state          := 0; // IDLE
            END_IF;
        ELSIF pendingConfirm AND doneSensor THEN
            // S10: Valve closed last scan, confirmed this scan
            IF fillsToday < 32767 THEN
                fillsToday := fillsToday + 1;
            END_IF;
            pendingConfirm := FALSE;
            state          := 0; // IDLE
        END_IF;
    END_IF;

    prevStartBtn  := startBtn;
    prevResetBtn  := resetBtn;
    prevValveOpen := valveOpen;
END_FUNCTION_BLOCK

(* ---- self-medium-04.raw_candidate_04.st ---- *)
FUNCTION_BLOCK FB
VAR_INPUT
    startBtn    : BOOL;
    resetBtn    : BOOL;
    doneSensor  : BOOL;
    targetVol   : REAL;
    flowVol     : REAL;
END_VAR
VAR_OUTPUT
    valveOpen   : BOOL := FALSE;
    fillsToday  : INT  := 0;
END_VAR
VAR
    state           : INT := 0; // 0=IDLE, 1=FILLING, 2=WAIT_CONFIRM
    accumulated     : REAL := 0.0;
    pendingConfirm  : BOOL := FALSE;
    prevStartBtn    : BOOL := FALSE;
    prevResetBtn    : BOOL := FALSE;
    prevValveOpen   : BOOL := FALSE;
    R_TRIG_reset    : R_TRIG;
    R_TRIG_start    : R_TRIG;
END_VAR
BEGIN
    (* ENGINEERING_CONTRACT
    ---------------------------------------------------------------------
    PUB001: Initialization - valve closed (valveOpen=FALSE), no pending
            confirmation (pendingConfirm=FALSE), fillsToday=0 on cold start.
    PUB002: Rising-edge detection for startBtn/resetBtn; pre-power state FALSE.
    PUB003: Scan execution order: reset(1)→start/new-bottle(2)→accumulate/
            close-on-target(3)→doneSensor read→confirm/count(4).
    PUB004: resetBtn rising edge has highest priority; clears all state,
            ignores same-scan start/flow/confirmation.
    PUB005: startBtn rising edge in IDLE/WAIT_CONFIRM starts new bottle,
            clears accumulation, opens valve. Prior pendingConfirm cancelled.
            New start during FILLING does NOT reset current bottle.
    PUB006: Accumulate flowVol every scan including startup scan.
    PUB007: When accumulated >= targetVol, close valve and set pendingConfirm
            immediately in same scan.
    PUB008: After closing, read doneSensor same scan. If TRUE, confirm/count
            immediately. If FALSE, wait for first TRUE (unless reset/new-start).
    PUB009: Each confirmation increments fillsToday by 1. At 32767, confirm
            completes but count stays at 32767.
    PUB010: Confirmation clears pendingConfirm. Continuous TRUE does not
            double-count. New-bottle start-cancel clears pendingConfirm.
    PUB011: fillsToday is INT; reset clears to 0.
    ---------------------------------------------------------------------
    OUTPUT RETENTION:
    - valveOpen: held open during FILLING until target met or reset/start.
    - fillsToday: monotonic non-decreasing except reset (S3); max 32767.
    - pendingConfirm: held TRUE from close until first TRUE doneSensor.
    EXPLICIT RESET: resetBtn rising edge clears accumulated, fillsToday,
            valveOpen, pendingConfirm, state→0(IDLE).
    SAME-SCAN PRIORITY: reset > close-on-target-with-confirm > start.
    UNITS/BOUNDARIES: accumulated REAL mL; fillsToday INT [0..32767];
            targetVol, flowVol REAL mL.
    ---------------------------------------------------------------------
    *)

    // Update edge detectors every scan
    R_TRIG_reset(CLK := resetBtn);
    R_TRIG_start(CLK := startBtn);

    // --- Step 1: Reset (highest priority) ---
    IF R_TRIG_reset.Q THEN
        accumulated    := 0.0;
        fillsToday     := 0;
        valveOpen      := FALSE;
        pendingConfirm := FALSE;
        state          := 0; // IDLE
        prevValveOpen  := FALSE;
        prevStartBtn   := startBtn;
        prevResetBtn   := resetBtn;
        RETURN;
    END_IF;

    // --- Step 2: Start new bottle ---
    IF R_TRIG_start.Q THEN
        IF state = 2 THEN // WAIT_CONFIRM
            pendingConfirm := FALSE;
        END_IF;
        IF state <> 1 THEN // not FILLING
            accumulated  := 0.0;
            valveOpen    := TRUE;
            state        := 1; // FILLING
        END_IF;
    END_IF;

    // --- Step 3: Accumulate and close on target ---
    IF state = 1 THEN // FILLING
        accumulated := accumulated + flowVol;
        IF accumulated >= targetVol THEN
            valveOpen      := FALSE;
            pendingConfirm := TRUE;
            state          := 2; // WAIT_CONFIRM
        END_IF;
    END_IF;

    // --- Step 4: Confirm/count on doneSensor ---
    IF pendingConfirm THEN
        IF doneSensor THEN
            IF fillsToday < 32767 THEN
                fillsToday := fillsToday + 1;
            END_IF;
            pendingConfirm := FALSE;
            state          := 0; // IDLE
        END_IF;
    END_IF;

    // Update previous states for edge detection
    prevStartBtn  := startBtn;
    prevResetBtn  := resetBtn;
    prevValveOpen := valveOpen;
END_FUNCTION_BLOCK

(* ---- self-medium-05.candidate_01.st ---- *)
FUNCTION_BLOCK FB
VAR_INPUT
    enable        : BOOL;
    resetBtn      : BOOL;
    scanSeconds   : LREAL;
    steamFlow     : LREAL;
    fuelFlow      : LREAL;
    steamTemp     : LREAL;
    steamPressure : LREAL;
END_VAR
VAR_OUTPUT
    qualified    : BOOL;
    dataFault    : BOOL;
    qualifiedTon : LREAL;
    fuelTon      : LREAL;
    revenue      : LREAL;
    cost         : LREAL;
    netProfit    : LREAL;
END_VAR
VAR
    prevResetBtn : BOOL := FALSE;
    localQualified : BOOL;
    localDataFault : BOOL;
    localResetRising : BOOL;
    tmpFuelIncrement : LREAL;
    tmpQualifiedIncrement : LREAL;
END_VAR
VAR_TEMP
    localSkipAccum : BOOL;
END_VAR
(*
ENGINEERING_CONTRACT
================================================================================
 PUB001: enable=TRUE → metering active; FALSE → hold accumulators (unless reset).
 PUB002: resetBtn rising edge → immediate zero-clear of qualifiedTon & fuelTon.
 PUB003: qualifiedTon, fuelTon accumulate in t (kg/s × s ÷ 1000); revenue=ton×280.
 PUB005: qualifiedTon increment requires qualified flag TRUE (see PUB001).
 PUB006: closed-interval qualification: temp∈[447,453] AND press∈[3750,3850].
 PUB007: fuelTon always accumulates when enable=TRUE AND no fault (independent of qualified).
 PUB008: dataFault when scanSeconds≤0 OR scanSeconds>10 OR flow out of [0,90]/[0,6].
 PUB009: reset rising edge PRIOR to fault freeze; both accumulators = 0.0 same-scan.
 PUB010: revenue/cost/netProfit update every scan (even when accumulation frozen).
 PUB011: qualifiedTon, fuelTon, revenue, cost ≥ 0 always; netProfit may be negative.
 PUB012: reset is edge-triggered (prevBtn memory); level-hold has no effect.
 PUB013–PUB016: scanSeconds, steamFlow, fuelFlow numeric bounds; fault gates accumulation.
================================================================================
Output states:
  qualified    | activation: steamTemp∈[447,453] ∧ steamPressure∈[3750,3850]; RETAINED via localQualified.
  dataFault    | activation: scanSeconds≤0 ∨ scanSeconds>10 ∨ steamFlow∉[0,90] ∨ fuelFlow∉[0,6]; RETAINED.
  qualifiedTon | hold_until_reset: cleared on resetBtn rising edge; no other reset.
  fuelTon      | hold_until_reset: cleared on resetBtn rising edge; no other reset.
  revenue/cost/netProfit | computed every scan from accumulator values; not independently latched.

Units/boundaries:
  scanSeconds: >0 (exclusive) and ≤10 (inclusive); unit s.
  steamFlow: [0,90] kg/s; fuelFlow: [0,6] kg/s.
  Conversion: kg/s × s ÷ 1000 = t.
  Prices: steam 280 元/t; fuel 1500 元/t.
================================================================================
*)
BEGIN
    (* Edge detection for reset (PUB012) *)
    localResetRising := resetBtn AND NOT prevResetBtn;

    (* Fault detection (PUB008) *)
    localDataFault := (scanSeconds <= 0.0) OR (scanSeconds > 10.0)
                      OR (steamFlow < 0.0) OR (steamFlow > 90.0)
                      OR (fuelFlow < 0.0) OR (fuelFlow > 6.0);

    (* Qualified flag — closed interval (PUB006) *)
    localQualified := (steamTemp >= 447.0) AND (steamTemp <= 453.0)
                      AND (steamPressure >= 3750.0) AND (steamPressure <= 3850.0);

    (* Accumulation: reset takes priority (PUB009, PUB002) *)
    IF localResetRising THEN
        qualifiedTon := 0.0;
        fuelTon      := 0.0;
        localSkipAccum := TRUE;
    ELSIF enable AND NOT localDataFault THEN
        (* PUB007: fuelTon increments regardless of qualified status *)
        tmpFuelIncrement := fuelFlow * scanSeconds / 1000.0;
        fuelTon := fuelTon + tmpFuelIncrement;

        (* PUB003, PUB005: qualifiedTon increments only when qualified=TRUE *)
        IF localQualified THEN
            tmpQualifiedIncrement := steamFlow * scanSeconds / 1000.0;
            qualifiedTon := qualifiedTon + tmpQualifiedIncrement;
        END_IF;

        localSkipAccum := FALSE;
    ELSE
        (* PUB009: fault or disabled without reset → hold accumulators *)
        localSkipAccum := FALSE;
    END_IF;

    (* Monetary calculations every scan (PUB010) *)
    revenue  := qualifiedTon * 280.0;
    cost     := fuelTon * 1500.0;
    netProfit := revenue - cost;

    (* Assign public outputs *)
    qualified    := localQualified;
    dataFault    := localDataFault;

    (* Update edge-detection memory for next scan (PUB012) *)
    prevResetBtn := resetBtn;
END_FUNCTION_BLOCK
(* CONTRACT_RULES [] *)

(* ---- self-medium-05.candidate_02.st ---- *)
FUNCTION_BLOCK FB
VAR_INPUT
    enable        : BOOL;
    resetBtn      : BOOL;
    scanSeconds   : LREAL;
    steamFlow     : LREAL;
    fuelFlow      : LREAL;
    steamTemp     : LREAL;
    steamPressure : LREAL;
END_VAR
VAR_OUTPUT
    qualified    : BOOL;
    dataFault    : BOOL;
    qualifiedTon : LREAL;
    fuelTon      : LREAL;
    revenue      : LREAL;
    cost         : LREAL;
    netProfit    : LREAL;
END_VAR
VAR
    prevResetBtn     : BOOL := FALSE;
    tmpResetRising   : BOOL;
    tmpDataFault     : BOOL;
    tmpQualified     : BOOL;
    tmpFuelIncrement : LREAL;
    tmpQualIncrement : LREAL;
END_VAR
(*
ENGINEERING_CONTRACT
================================================================================
 PUB001: enable=TRUE → metering active; FALSE → hold accumulators (unless reset).
 PUB002: resetBtn rising edge → immediate zero-clear of qualifiedTon & fuelTon.
 PUB003: qualifiedTon, fuelTon accumulate in t (kg/s × s ÷ 1000); revenue=ton×280.
 PUB005: qualifiedTon increment requires qualified flag TRUE (see PUB001).
 PUB006: closed-interval qualification: temp∈[447,453] AND press∈[3750,3850].
 PUB007: fuelTon always accumulates when enable=TRUE AND no fault (independent of qualified).
 PUB008: dataFault when scanSeconds≤0 OR scanSeconds>10 OR flow out of [0,90]/[0,6].
 PUB009: reset rising edge PRIOR to fault freeze; both accumulators = 0.0 same-scan.
 PUB010: revenue/cost/netProfit update every scan (even when accumulation frozen).
 PUB011: qualifiedTon, fuelTon, revenue, cost ≥ 0 always; netProfit may be negative.
 PUB012: reset is edge-triggered (prevBtn memory); level-hold has no effect.
 PUB013–PUB016: scanSeconds, steamFlow, fuelFlow numeric bounds; fault gates accumulation.
================================================================================
Output states:
  qualified    | activation: steamTemp∈[447,453] ∧ steamPressure∈[3750,3850]; RETAINED.
  dataFault    | activation: scanSeconds≤0 ∨ scanSeconds>10 ∨ steamFlow∉[0,90] ∨ fuelFlow∉[0,6]; RETAINED.
  qualifiedTon | hold_until_reset: cleared on resetBtn rising edge; no other reset.
  fuelTon      | hold_until_reset: cleared on resetBtn rising edge; no other reset.
  revenue/cost/netProfit | computed every scan from accumulator values; not independently latched.
================================================================================
*)
BEGIN
    tmpResetRising := resetBtn AND NOT prevResetBtn;
    tmpDataFault := (scanSeconds <= 0.0) OR (scanSeconds > 10.0)
                    OR (steamFlow < 0.0) OR (steamFlow > 90.0)
                    OR (fuelFlow < 0.0) OR (fuelFlow > 6.0);
    tmpQualified := (steamTemp >= 447.0) AND (steamTemp <= 453.0)
                    AND (steamPressure >= 3750.0) AND (steamPressure <= 3850.0);

    IF tmpResetRising THEN
        qualifiedTon := 0.0;
        fuelTon := 0.0;
    ELSIF enable AND NOT tmpDataFault THEN
        tmpFuelIncrement := fuelFlow * scanSeconds / 1000.0;
        fuelTon := fuelTon + tmpFuelIncrement;
        IF tmpQualified THEN
            tmpQualIncrement := steamFlow * scanSeconds / 1000.0;
            qualifiedTon := qualifiedTon + tmpQualIncrement;
        END_IF;
    END_IF;

    revenue := qualifiedTon * 280.0;
    cost := fuelTon * 1500.0;
    netProfit := revenue - cost;

    qualified := tmpQualified;
    dataFault := tmpDataFault;

    prevResetBtn := resetBtn;
END_FUNCTION_BLOCK
(* CONTRACT_RULES [] *)

(* ---- self-medium-05.candidate_03.st ---- *)
FUNCTION_BLOCK FB
VAR_INPUT
    enable        : BOOL;
    resetBtn      : BOOL;
    scanSeconds   : LREAL;
    steamFlow     : LREAL;
    fuelFlow      : LREAL;
    steamTemp     : LREAL;
    steamPressure : LREAL;
END_VAR
VAR_OUTPUT
    qualified    : BOOL;
    dataFault    : BOOL;
    qualifiedTon : LREAL;
    fuelTon      : LREAL;
    revenue      : LREAL;
    cost         : LREAL;
    netProfit    : LREAL;
END_VAR
VAR
    prevResetBtn     : BOOL := FALSE;
    tmpQualified     : BOOL;
    tmpDataFault     : BOOL;
    tmpResetRising   : BOOL;
    tmpFuelInc       : LREAL;
    tmpQualInc       : LREAL;
END_VAR
(*
ENGINEERING_CONTRACT
================================================================================
 PUB001: enable=TRUE → metering active; FALSE → hold accumulators (unless reset).
 PUB002: resetBtn rising edge → immediate zero-clear of qualifiedTon & fuelTon.
 PUB003: qualifiedTon, fuelTon accumulate in t (kg/s × s ÷ 1000); revenue=ton×280.
 PUB005: qualifiedTon increment requires qualified flag TRUE (see PUB001).
 PUB006: closed-interval qualification: temp∈[447,453] AND press∈[3750,3850].
 PUB007: fuelTon always accumulates when enable=TRUE AND no fault (independent of qualified).
 PUB008: dataFault when scanSeconds≤0 OR scanSeconds>10 OR flow out of [0,90]/[0,6].
 PUB009: reset rising edge PRIOR to fault freeze; both accumulators = 0.0 same-scan.
 PUB010: revenue/cost/netProfit update every scan (even when accumulation frozen).
 PUB011: qualifiedTon, fuelTon, revenue, cost ≥ 0 always; netProfit may be negative.
 PUB012: reset is edge-triggered (prevBtn memory); level-hold has no effect.
 PUB013–PUB016: scanSeconds, steamFlow, fuelFlow numeric bounds; fault gates accumulation.
================================================================================
Output states:
  qualified    | activation: steamTemp∈[447,453] ∧ steamPressure∈[3750,3850]; RETAINED.
  dataFault    | activation: scanSeconds≤0 ∨ scanSeconds>10 ∨ steamFlow∉[0,90] ∨ fuelFlow∉[0,6]; RETAINED.
  qualifiedTon | hold_until_reset: cleared on resetBtn rising edge; no other reset.
  fuelTon      | hold_until_reset: cleared on resetBtn rising edge; no other reset.
  revenue/cost/netProfit | computed every scan from accumulator values; not independently latched.
================================================================================
*)
BEGIN
    tmpResetRising := resetBtn AND NOT prevResetBtn;

    tmpDataFault := (scanSeconds <= 0.0) OR (scanSeconds > 10.0)
                    OR (steamFlow < 0.0) OR (steamFlow > 90.0)
                    OR (fuelFlow < 0.0) OR (fuelFlow > 6.0);

    tmpQualified := (steamTemp >= 447.0) AND (steamTemp <= 453.0)
                    AND (steamPressure >= 3750.0) AND (steamPressure <= 3850.0);

    IF tmpResetRising THEN
        qualifiedTon := 0.0;
        fuelTon := 0.0;
    ELSIF enable AND NOT tmpDataFault THEN
        tmpFuelInc := fuelFlow * scanSeconds / 1000.0;
        fuelTon := fuelTon + tmpFuelInc;
        IF tmpQualified THEN
            tmpQualInc := steamFlow * scanSeconds / 1000.0;
            qualifiedTon := qualifiedTon + tmpQualInc;
        END_IF;
    END_IF;

    revenue := qualifiedTon * 280.0;
    cost := fuelTon * 1500.0;
    netProfit := revenue - cost;

    qualified := tmpQualified;
    dataFault := tmpDataFault;

    prevResetBtn := resetBtn;
END_FUNCTION_BLOCK
(* CONTRACT_RULES [] *)

(* ---- self-medium-05.candidate_04.st ---- *)
FUNCTION_BLOCK FB
VAR_INPUT
    enable        : BOOL;
    resetBtn      : BOOL;
    scanSeconds   : LREAL;
    steamFlow     : LREAL;
    fuelFlow      : LREAL;
    steamTemp     : LREAL;
    steamPressure : LREAL;
END_VAR
VAR_OUTPUT
    qualified    : BOOL;
    dataFault    : BOOL;
    qualifiedTon : LREAL;
    fuelTon      : LREAL;
    revenue      : LREAL;
    cost         : LREAL;
    netProfit    : LREAL;
END_VAR
VAR
    prevResetBtn      : BOOL := FALSE;
    localResetRising  : BOOL;
    localDataFault    : BOOL;
    localQualified    : BOOL;
    tmpFuelInc        : LREAL;
    tmpQualInc        : LREAL;
END_VAR
(*
ENGINEERING_CONTRACT
================================================================================
 PUB001: enable=TRUE → metering active; FALSE → hold accumulators (unless reset).
 PUB002: resetBtn rising edge → immediate zero-clear of qualifiedTon & fuelTon.
 PUB003: qualifiedTon, fuelTon accumulate in t (kg/s × s ÷ 1000); revenue=ton×280.
 PUB005: qualifiedTon increment requires qualified flag TRUE (see PUB001).
 PUB006: closed-interval qualification: temp∈[447,453] AND press∈[3750,3850].
 PUB007: fuelTon always accumulates when enable=TRUE AND no fault (independent of qualified).
 PUB008: dataFault when scanSeconds≤0 OR scanSeconds>10 OR flow out of [0,90]/[0,6].
 PUB009: reset rising edge PRIOR to fault freeze; both accumulators = 0.0 same-scan.
 PUB010: revenue/cost/netProfit update every scan (even when accumulation frozen).
 PUB011: qualifiedTon, fuelTon, revenue, cost ≥ 0 always; netProfit may be negative.
 PUB012: reset is edge-triggered (prevBtn memory); level-hold has no effect.
 PUB013–PUB016: scanSeconds, steamFlow, fuelFlow numeric bounds; fault gates accumulation.
================================================================================
Output states:
  qualified    | activation: steamTemp∈[447,453] ∧ steamPressure∈[3750,3850]; RETAINED.
  dataFault    | activation: scanSeconds≤0 ∨ scanSeconds>10 ∨ steamFlow∉[0,90] ∨ fuelFlow∉[0,6]; RETAINED.
  qualifiedTon | hold_until_reset: cleared on resetBtn rising edge; no other reset.
  fuelTon      | hold_until_reset: cleared on resetBtn rising edge; no other reset.
  revenue/cost/netProfit | computed every scan from accumulator values; not independently latched.
Units/boundaries:
  scanSeconds: >0 (exclusive) and ≤10 (inclusive); unit s.
  steamFlow: [0,90] kg/s; fuelFlow: [0,6] kg/s.
  Conversion: kg/s × s ÷ 1000 = t.
  Prices: steam 280 元/t; fuel 1500 元/t.
================================================================================
*)
BEGIN
    (* Edge detection for reset (PUB012) *)
    localResetRising := resetBtn AND NOT prevResetBtn;

    (* Fault detection (PUB008) *)
    localDataFault := (scanSeconds <= 0.0) OR (scanSeconds > 10.0)
                      OR (steamFlow < 0.0) OR (steamFlow > 90.0)
                      OR (fuelFlow < 0.0) OR (fuelFlow > 6.0);

    (* Qualified flag — closed interval (PUB006) *)
    localQualified := (steamTemp >= 447.0) AND (steamTemp <= 453.0)
                      AND (steamPressure >= 3750.0) AND (steamPressure <= 3850.0);

    (* Accumulation: reset takes priority (PUB009, PUB002) *)
    IF localResetRising THEN
        qualifiedTon := 0.0;
        fuelTon      := 0.0;
    ELSIF enable AND NOT localDataFault THEN
        (* PUB007: fuelTon increments regardless of qualified status *)
        tmpFuelInc := fuelFlow * scanSeconds / 1000.0;
        fuelTon := fuelTon + tmpFuelInc;

        (* PUB003, PUB005: qualifiedTon increments only when qualified=TRUE *)
        IF localQualified THEN
            tmpQualInc := steamFlow * scanSeconds / 1000.0;
            qualifiedTon := qualifiedTon + tmpQualInc;
        END_IF;
    END_IF;

    (* Monetary calculations every scan (PUB010) *)
    revenue   := qualifiedTon * 280.0;
    cost      := fuelTon * 1500.0;
    netProfit := revenue - cost;

    (* Assign public outputs *)
    qualified    := localQualified;
    dataFault    := localDataFault;

    (* Update edge-detection memory for next scan (PUB012) *)
    prevResetBtn := resetBtn;
END_FUNCTION_BLOCK
(* CONTRACT_RULES [] *)

(* ---- self-medium-05.raw_candidate_01.st ---- *)
FUNCTION_BLOCK FB
VAR_INPUT
    enable        : BOOL;
    resetBtn      : BOOL;
    scanSeconds   : LREAL;
    steamFlow     : LREAL;
    fuelFlow      : LREAL;
    steamTemp     : LREAL;
    steamPressure : LREAL;
END_VAR
VAR_OUTPUT
    qualified    : BOOL;
    dataFault    : BOOL;
    qualifiedTon : LREAL;
    fuelTon      : LREAL;
    revenue      : LREAL;
    cost         : LREAL;
    netProfit    : LREAL;
END_VAR
VAR
    prevResetBtn : BOOL := FALSE;
    localQualified : BOOL;
    localDataFault : BOOL;
    localResetRising : BOOL;
    tmpFuelIncrement : LREAL;
    tmpQualifiedIncrement : LREAL;
END_VAR
VAR_TEMP
    localSkipAccum : BOOL;
END_VAR
(*
ENGINEERING_CONTRACT
================================================================================
 PUB001: enable=TRUE → metering active; FALSE → hold accumulators (unless reset).
 PUB002: resetBtn rising edge → immediate zero-clear of qualifiedTon & fuelTon.
 PUB003: qualifiedTon, fuelTon accumulate in t (kg/s × s ÷ 1000); revenue=ton×280.
 PUB005: qualifiedTon increment requires qualified flag TRUE (see PUB001).
 PUB006: closed-interval qualification: temp∈[447,453] AND press∈[3750,3850].
 PUB007: fuelTon always accumulates when enable=TRUE AND no fault (independent of qualified).
 PUB008: dataFault when scanSeconds≤0 OR scanSeconds>10 OR flow out of [0,90]/[0,6].
 PUB009: reset rising edge PRIOR to fault freeze; both accumulators = 0.0 same-scan.
 PUB010: revenue/cost/netProfit update every scan (even when accumulation frozen).
 PUB011: qualifiedTon, fuelTon, revenue, cost ≥ 0 always; netProfit may be negative.
 PUB012: reset is edge-triggered (prevBtn memory); level-hold has no effect.
 PUB013–PUB016: scanSeconds, steamFlow, fuelFlow numeric bounds; fault gates accumulation.
================================================================================
Output states:
  qualified    | activation: steamTemp∈[447,453] ∧ steamPressure∈[3750,3850]; RETAINED via localQualified.
  dataFault    | activation: scanSeconds≤0 ∨ scanSeconds>10 ∨ steamFlow∉[0,90] ∨ fuelFlow∉[0,6]; RETAINED.
  qualifiedTon | hold_until_reset: cleared on resetBtn rising edge; no other reset.
  fuelTon      | hold_until_reset: cleared on resetBtn rising edge; no other reset.
  revenue/cost/netProfit | computed every scan from accumulator values; not independently latched.

Units/boundaries:
  scanSeconds: >0 (exclusive) and ≤10 (inclusive); unit s.
  steamFlow: [0,90] kg/s; fuelFlow: [0,6] kg/s.
  Conversion: kg/s × s ÷ 1000 = t.
  Prices: steam 280 元/t; fuel 1500 元/t.
================================================================================
*)
BEGIN
    (* Edge detection for reset (PUB012) *)
    localResetRising := resetBtn AND NOT prevResetBtn;

    (* Fault detection (PUB008) *)
    localDataFault := (scanSeconds <= 0.0) OR (scanSeconds > 10.0)
                      OR (steamFlow < 0.0) OR (steamFlow > 90.0)
                      OR (fuelFlow < 0.0) OR (fuelFlow > 6.0);

    (* Qualified flag — closed interval (PUB006) *)
    localQualified := (steamTemp >= 447.0) AND (steamTemp <= 453.0)
                      AND (steamPressure >= 3750.0) AND (steamPressure <= 3850.0);

    (* Accumulation: reset takes priority (PUB009, PUB002) *)
    IF localResetRising THEN
        qualifiedTon := 0.0;
        fuelTon      := 0.0;
        localSkipAccum := TRUE;
    ELSIF enable AND NOT localDataFault THEN
        (* PUB007: fuelTon increments regardless of qualified status *)
        tmpFuelIncrement := fuelFlow * scanSeconds / 1000.0;
        fuelTon := fuelTon + tmpFuelIncrement;

        (* PUB003, PUB005: qualifiedTon increments only when qualified=TRUE *)
        IF localQualified THEN
            tmpQualifiedIncrement := steamFlow * scanSeconds / 1000.0;
            qualifiedTon := qualifiedTon + tmpQualifiedIncrement;
        END_IF;

        localSkipAccum := FALSE;
    ELSE
        (* PUB009: fault or disabled without reset → hold accumulators *)
        localSkipAccum := FALSE;
    END_IF;

    (* Monetary calculations every scan (PUB010) *)
    revenue  := qualifiedTon * 280.0;
    cost     := fuelTon * 1500.0;
    netProfit := revenue - cost;

    (* Assign public outputs *)
    qualified    := localQualified;
    dataFault    := localDataFault;

    (* Update edge-detection memory for next scan (PUB012) *)
    prevResetBtn := resetBtn;
END_FUNCTION_BLOCK
(* CONTRACT_RULES [] *)

(* ---- self-medium-05.raw_candidate_02.st ---- *)
FUNCTION_BLOCK FB
VAR_INPUT
    enable        : BOOL;
    resetBtn      : BOOL;
    scanSeconds   : LREAL;
    steamFlow     : LREAL;
    fuelFlow      : LREAL;
    steamTemp     : LREAL;
    steamPressure : LREAL;
END_VAR
VAR_OUTPUT
    qualified    : BOOL;
    dataFault    : BOOL;
    qualifiedTon : LREAL;
    fuelTon      : LREAL;
    revenue      : LREAL;
    cost         : LREAL;
    netProfit    : LREAL;
END_VAR
VAR
    prevResetBtn     : BOOL := FALSE;
    tmpResetRising   : BOOL;
    tmpDataFault     : BOOL;
    tmpQualified     : BOOL;
    tmpFuelIncrement : LREAL;
    tmpQualIncrement : LREAL;
END_VAR
(*
ENGINEERING_CONTRACT
================================================================================
 PUB001: enable=TRUE → metering active; FALSE → hold accumulators (unless reset).
 PUB002: resetBtn rising edge → immediate zero-clear of qualifiedTon & fuelTon.
 PUB003: qualifiedTon, fuelTon accumulate in t (kg/s × s ÷ 1000); revenue=ton×280.
 PUB005: qualifiedTon increment requires qualified flag TRUE (see PUB001).
 PUB006: closed-interval qualification: temp∈[447,453] AND press∈[3750,3850].
 PUB007: fuelTon always accumulates when enable=TRUE AND no fault (independent of qualified).
 PUB008: dataFault when scanSeconds≤0 OR scanSeconds>10 OR flow out of [0,90]/[0,6].
 PUB009: reset rising edge PRIOR to fault freeze; both accumulators = 0.0 same-scan.
 PUB010: revenue/cost/netProfit update every scan (even when accumulation frozen).
 PUB011: qualifiedTon, fuelTon, revenue, cost ≥ 0 always; netProfit may be negative.
 PUB012: reset is edge-triggered (prevBtn memory); level-hold has no effect.
 PUB013–PUB016: scanSeconds, steamFlow, fuelFlow numeric bounds; fault gates accumulation.
================================================================================
Output states:
  qualified    | activation: steamTemp∈[447,453] ∧ steamPressure∈[3750,3850]; RETAINED.
  dataFault    | activation: scanSeconds≤0 ∨ scanSeconds>10 ∨ steamFlow∉[0,90] ∨ fuelFlow∉[0,6]; RETAINED.
  qualifiedTon | hold_until_reset: cleared on resetBtn rising edge; no other reset.
  fuelTon      | hold_until_reset: cleared on resetBtn rising edge; no other reset.
  revenue/cost/netProfit | computed every scan from accumulator values; not independently latched.
================================================================================
*)
BEGIN
    tmpResetRising := resetBtn AND NOT prevResetBtn;
    tmpDataFault := (scanSeconds <= 0.0) OR (scanSeconds > 10.0)
                    OR (steamFlow < 0.0) OR (steamFlow > 90.0)
                    OR (fuelFlow < 0.0) OR (fuelFlow > 6.0);
    tmpQualified := (steamTemp >= 447.0) AND (steamTemp <= 453.0)
                    AND (steamPressure >= 3750.0) AND (steamPressure <= 3850.0);

    IF tmpResetRising THEN
        qualifiedTon := 0.0;
        fuelTon := 0.0;
    ELSIF enable AND NOT tmpDataFault THEN
        tmpFuelIncrement := fuelFlow * scanSeconds / 1000.0;
        fuelTon := fuelTon + tmpFuelIncrement;
        IF tmpQualified THEN
            tmpQualIncrement := steamFlow * scanSeconds / 1000.0;
            qualifiedTon := qualifiedTon + tmpQualIncrement;
        END_IF;
    END_IF;

    revenue := qualifiedTon * 280.0;
    cost := fuelTon * 1500.0;
    netProfit := revenue - cost;

    qualified := tmpQualified;
    dataFault := tmpDataFault;

    prevResetBtn := resetBtn;
END_FUNCTION_BLOCK
(* CONTRACT_RULES [] *)

(* ---- self-medium-05.raw_candidate_03.st ---- *)
FUNCTION_BLOCK FB
VAR_INPUT
    enable        : BOOL;
    resetBtn      : BOOL;
    scanSeconds   : LREAL;
    steamFlow     : LREAL;
    fuelFlow      : LREAL;
    steamTemp     : LREAL;
    steamPressure : LREAL;
END_VAR
VAR_OUTPUT
    qualified    : BOOL;
    dataFault    : BOOL;
    qualifiedTon : LREAL;
    fuelTon      : LREAL;
    revenue      : LREAL;
    cost         : LREAL;
    netProfit    : LREAL;
END_VAR
VAR
    prevResetBtn     : BOOL := FALSE;
    tmpQualified     : BOOL;
    tmpDataFault     : BOOL;
    tmpResetRising   : BOOL;
    tmpFuelInc       : LREAL;
    tmpQualInc       : LREAL;
END_VAR
(*
ENGINEERING_CONTRACT
================================================================================
 PUB001: enable=TRUE → metering active; FALSE → hold accumulators (unless reset).
 PUB002: resetBtn rising edge → immediate zero-clear of qualifiedTon & fuelTon.
 PUB003: qualifiedTon, fuelTon accumulate in t (kg/s × s ÷ 1000); revenue=ton×280.
 PUB005: qualifiedTon increment requires qualified flag TRUE (see PUB001).
 PUB006: closed-interval qualification: temp∈[447,453] AND press∈[3750,3850].
 PUB007: fuelTon always accumulates when enable=TRUE AND no fault (independent of qualified).
 PUB008: dataFault when scanSeconds≤0 OR scanSeconds>10 OR flow out of [0,90]/[0,6].
 PUB009: reset rising edge PRIOR to fault freeze; both accumulators = 0.0 same-scan.
 PUB010: revenue/cost/netProfit update every scan (even when accumulation frozen).
 PUB011: qualifiedTon, fuelTon, revenue, cost ≥ 0 always; netProfit may be negative.
 PUB012: reset is edge-triggered (prevBtn memory); level-hold has no effect.
 PUB013–PUB016: scanSeconds, steamFlow, fuelFlow numeric bounds; fault gates accumulation.
================================================================================
Output states:
  qualified    | activation: steamTemp∈[447,453] ∧ steamPressure∈[3750,3850]; RETAINED.
  dataFault    | activation: scanSeconds≤0 ∨ scanSeconds>10 ∨ steamFlow∉[0,90] ∨ fuelFlow∉[0,6]; RETAINED.
  qualifiedTon | hold_until_reset: cleared on resetBtn rising edge; no other reset.
  fuelTon      | hold_until_reset: cleared on resetBtn rising edge; no other reset.
  revenue/cost/netProfit | computed every scan from accumulator values; not independently latched.
================================================================================
*)
BEGIN
    tmpResetRising := resetBtn AND NOT prevResetBtn;

    tmpDataFault := (scanSeconds <= 0.0) OR (scanSeconds > 10.0)
                    OR (steamFlow < 0.0) OR (steamFlow > 90.0)
                    OR (fuelFlow < 0.0) OR (fuelFlow > 6.0);

    tmpQualified := (steamTemp >= 447.0) AND (steamTemp <= 453.0)
                    AND (steamPressure >= 3750.0) AND (steamPressure <= 3850.0);

    IF tmpResetRising THEN
        qualifiedTon := 0.0;
        fuelTon := 0.0;
    ELSIF enable AND NOT tmpDataFault THEN
        tmpFuelInc := fuelFlow * scanSeconds / 1000.0;
        fuelTon := fuelTon + tmpFuelInc;
        IF tmpQualified THEN
            tmpQualInc := steamFlow * scanSeconds / 1000.0;
            qualifiedTon := qualifiedTon + tmpQualInc;
        END_IF;
    END_IF;

    revenue := qualifiedTon * 280.0;
    cost := fuelTon * 1500.0;
    netProfit := revenue - cost;

    qualified := tmpQualified;
    dataFault := tmpDataFault;

    prevResetBtn := resetBtn;
END_FUNCTION_BLOCK
(* CONTRACT_RULES [] *)

(* ---- self-medium-05.raw_candidate_04.st ---- *)
FUNCTION_BLOCK FB
VAR_INPUT
    enable        : BOOL;
    resetBtn      : BOOL;
    scanSeconds   : LREAL;
    steamFlow     : LREAL;
    fuelFlow      : LREAL;
    steamTemp     : LREAL;
    steamPressure : LREAL;
END_VAR
VAR_OUTPUT
    qualified    : BOOL;
    dataFault    : BOOL;
    qualifiedTon : LREAL;
    fuelTon      : LREAL;
    revenue      : LREAL;
    cost         : LREAL;
    netProfit    : LREAL;
END_VAR
VAR
    prevResetBtn      : BOOL := FALSE;
    localResetRising  : BOOL;
    localDataFault    : BOOL;
    localQualified    : BOOL;
    tmpFuelInc        : LREAL;
    tmpQualInc        : LREAL;
END_VAR
(*
ENGINEERING_CONTRACT
================================================================================
 PUB001: enable=TRUE → metering active; FALSE → hold accumulators (unless reset).
 PUB002: resetBtn rising edge → immediate zero-clear of qualifiedTon & fuelTon.
 PUB003: qualifiedTon, fuelTon accumulate in t (kg/s × s ÷ 1000); revenue=ton×280.
 PUB005: qualifiedTon increment requires qualified flag TRUE (see PUB001).
 PUB006: closed-interval qualification: temp∈[447,453] AND press∈[3750,3850].
 PUB007: fuelTon always accumulates when enable=TRUE AND no fault (independent of qualified).
 PUB008: dataFault when scanSeconds≤0 OR scanSeconds>10 OR flow out of [0,90]/[0,6].
 PUB009: reset rising edge PRIOR to fault freeze; both accumulators = 0.0 same-scan.
 PUB010: revenue/cost/netProfit update every scan (even when accumulation frozen).
 PUB011: qualifiedTon, fuelTon, revenue, cost ≥ 0 always; netProfit may be negative.
 PUB012: reset is edge-triggered (prevBtn memory); level-hold has no effect.
 PUB013–PUB016: scanSeconds, steamFlow, fuelFlow numeric bounds; fault gates accumulation.
================================================================================
Output states:
  qualified    | activation: steamTemp∈[447,453] ∧ steamPressure∈[3750,3850]; RETAINED.
  dataFault    | activation: scanSeconds≤0 ∨ scanSeconds>10 ∨ steamFlow∉[0,90] ∨ fuelFlow∉[0,6]; RETAINED.
  qualifiedTon | hold_until_reset: cleared on resetBtn rising edge; no other reset.
  fuelTon      | hold_until_reset: cleared on resetBtn rising edge; no other reset.
  revenue/cost/netProfit | computed every scan from accumulator values; not independently latched.
Units/boundaries:
  scanSeconds: >0 (exclusive) and ≤10 (inclusive); unit s.
  steamFlow: [0,90] kg/s; fuelFlow: [0,6] kg/s.
  Conversion: kg/s × s ÷ 1000 = t.
  Prices: steam 280 元/t; fuel 1500 元/t.
================================================================================
*)
BEGIN
    (* Edge detection for reset (PUB012) *)
    localResetRising := resetBtn AND NOT prevResetBtn;

    (* Fault detection (PUB008) *)
    localDataFault := (scanSeconds <= 0.0) OR (scanSeconds > 10.0)
                      OR (steamFlow < 0.0) OR (steamFlow > 90.0)
                      OR (fuelFlow < 0.0) OR (fuelFlow > 6.0);

    (* Qualified flag — closed interval (PUB006) *)
    localQualified := (steamTemp >= 447.0) AND (steamTemp <= 453.0)
                      AND (steamPressure >= 3750.0) AND (steamPressure <= 3850.0);

    (* Accumulation: reset takes priority (PUB009, PUB002) *)
    IF localResetRising THEN
        qualifiedTon := 0.0;
        fuelTon      := 0.0;
    ELSIF enable AND NOT localDataFault THEN
        (* PUB007: fuelTon increments regardless of qualified status *)
        tmpFuelInc := fuelFlow * scanSeconds / 1000.0;
        fuelTon := fuelTon + tmpFuelInc;

        (* PUB003, PUB005: qualifiedTon increments only when qualified=TRUE *)
        IF localQualified THEN
            tmpQualInc := steamFlow * scanSeconds / 1000.0;
            qualifiedTon := qualifiedTon + tmpQualInc;
        END_IF;
    END_IF;

    (* Monetary calculations every scan (PUB010) *)
    revenue   := qualifiedTon * 280.0;
    cost      := fuelTon * 1500.0;
    netProfit := revenue - cost;

    (* Assign public outputs *)
    qualified    := localQualified;
    dataFault    := localDataFault;

    (* Update edge-detection memory for next scan (PUB012) *)
    prevResetBtn := resetBtn;
END_FUNCTION_BLOCK
(* CONTRACT_RULES [] *)
